  movel([-0.121105, -0.780827, -2.794142, -1.137419, 1.570796, 1.449692],accel_mss,speed_ms,0,blend_radius_m)
  movel([-0.120159, -0.781005, -2.794114, -1.137271, 1.570796, 1.450637],accel_mss,speed_ms,0,blend_radius_m)
  movel([-0.119008, -0.782524, -2.793869, -1.135997, 1.570796, 1.451789],accel_mss,speed_ms,0,blend_radius_m)
  movel([-0.118135, -0.785303, -2.793417, -1.133668, 1.570796, 1.452661],accel_mss,speed_ms,0,blend_radius_m)
  movel([-0.117601, -0.788380, -2.792913, -1.131096, 1.570796, 1.453195],accel_mss,speed_ms,0,blend_radius_m)
  movel([-0.115239, -0.783750, -2.793670, -1.134969, 1.570796, 1.455558],accel_mss,speed_ms,0,blend_radius_m)
  movel([-0.112520, -0.779061, -2.794425, -1.138903, 1.570796, 1.458276],accel_mss,speed_ms,0,blend_radius_m)
  movel([-0.109499, -0.774375, -2.795169, -1.142845, 1.570796, 1.461298],accel_mss,speed_ms,0,blend_radius_m)
  movel([-0.106241, -0.769762, -2.795890, -1.146737, 1.570796, 1.464556],accel_mss,speed_ms,0,blend_radius_m)
  movel([-0.099689, -0.760491, -2.797308, -1.154590, 1.570796, 1.471108],accel_mss,speed_ms,0,blend_radius_m)
  movel([-0.097728, -0.757937, -2.797692, -1.156760, 1.570796, 1.473068],accel_mss,speed_ms,0,blend_radius_m)
  movel([-0.095794, -0.755653, -2.798032, -1.158704, 1.570796, 1.475003],accel_mss,speed_ms,0,blend_radius_m)
  movel([-0.093954, -0.753818, -2.798303, -1.160268, 1.570796, 1.476842],accel_mss,speed_ms,0,blend_radius_m)
  movel([-0.092299, -0.752614, -2.798480, -1.161295, 1.570796, 1.478498],accel_mss,speed_ms,0,blend_radius_m)
  movel([-0.090884, -0.752253, -2.798533, -1.161603, 1.570796, 1.479912],accel_mss,speed_ms,0,blend_radius_m)
  movel([-0.089878, -0.752769, -2.798457, -1.161162, 1.570796, 1.480919],accel_mss,speed_ms,0,blend_radius_m)
  movel([-0.089251, -0.753972, -2.798280, -1.160137, 1.570796, 1.481545],accel_mss,speed_ms,0,blend_radius_m)
  movel([-0.088991, -0.755673, -2.798029, -1.158687, 1.570796, 1.481805],accel_mss,speed_ms,0,blend_radius_m)
  movel([-0.089073, -0.757680, -2.797730, -1.156979, 1.570796, 1.481724],accel_mss,speed_ms,0,blend_radius_m)
  movel([-0.089471, -0.759797, -2.797413, -1.155179, 1.570796, 1.481326],accel_mss,speed_ms,0,blend_radius_m)
  movel([-0.090165, -0.761839, -2.797105, -1.153445, 1.570796, 1.480631],accel_mss,speed_ms,0,blend_radius_m)
  movel([-0.091138, -0.763618, -2.796835, -1.151936, 1.570796, 1.479658],accel_mss,speed_ms,0,blend_radius_m)
  movel([-0.085055, -0.755408, -2.798068, -1.158913, 1.570796, 1.485742],accel_mss,speed_ms,0,blend_radius_m)
  movel([-0.081792, -0.751409, -2.798657, -1.162323, 1.570796, 1.489004],accel_mss,speed_ms,0,blend_radius_m)
  movel([-0.078396, -0.747530, -2.799220, -1.165639, 1.570796, 1.492400],accel_mss,speed_ms,0,blend_radius_m)
  movel([-0.074888, -0.743806, -2.799755, -1.168828, 1.570796, 1.495909],accel_mss,speed_ms,0,blend_radius_m)
  movel([-0.071275, -0.740275, -2.800255, -1.171859, 1.570796, 1.499521],accel_mss,speed_ms,0,blend_radius_m)
  movel([-0.067576, -0.736976, -2.800718, -1.174695, 1.570796, 1.503221],accel_mss,speed_ms,0,blend_radius_m)
  movel([-0.063806, -0.733944, -2.801138, -1.177307, 1.570796, 1.506991],accel_mss,speed_ms,0,blend_radius_m)
  movel([-0.061242, -0.732398, -2.801351, -1.178640, 1.570796, 1.509554],accel_mss,speed_ms,0,blend_radius_m)
  movel([-0.058496, -0.731434, -2.801483, -1.179472, 1.570796, 1.512301],accel_mss,speed_ms,0,blend_radius_m)
  movel([-0.057304, -0.731323, -2.801498, -1.179568, 1.570796, 1.513493],accel_mss,speed_ms,0,blend_radius_m)
  movel([-0.056360, -0.731534, -2.801469, -1.179386, 1.570796, 1.514437],accel_mss,speed_ms,0,blend_radius_m)
  movel([-0.055759, -0.732128, -2.801388, -1.178873, 1.570796, 1.515037],accel_mss,speed_ms,0,blend_radius_m)
  movel([-0.055607, -0.733168, -2.801245, -1.177976, 1.570796, 1.515190],accel_mss,speed_ms,0,blend_radius_m)
  movel([-0.055970, -0.734525, -2.801058, -1.176806, 1.570796, 1.514827],accel_mss,speed_ms,0,blend_radius_m)
  movel([-0.056714, -0.736045, -2.800847, -1.175497, 1.570796, 1.514083],accel_mss,speed_ms,0,blend_radius_m)
  movel([-0.058927, -0.739452, -2.800371, -1.172566, 1.570796, 1.511869],accel_mss,speed_ms,0,blend_radius_m)
  movel([-0.061573, -0.742637, -2.799921, -1.169831, 1.570796, 1.509223],accel_mss,speed_ms,0,blend_radius_m)
  movel([-0.064470, -0.745574, -2.799502, -1.167314, 1.570796, 1.506326],accel_mss,speed_ms,0,blend_radius_m)
  movel([-0.067437, -0.748234, -2.799119, -1.165036, 1.570796, 1.503359],accel_mss,speed_ms,0,blend_radius_m)
  movel([-0.063607, -0.746740, -2.799334, -1.166315, 1.570796, 1.507189],accel_mss,speed_ms,0,blend_radius_m)
  movel([-0.059620, -0.744795, -2.799614, -1.167981, 1.570796, 1.511176],accel_mss,speed_ms,0,blend_radius_m)
  movel([-0.055519, -0.742424, -2.799951, -1.170014, 1.570796, 1.515278],accel_mss,speed_ms,0,blend_radius_m)
  movel([-0.051338, -0.739647, -2.800344, -1.172398, 1.570796, 1.519459],accel_mss,speed_ms,0,blend_radius_m)
  movel([-0.048030, -0.737110, -2.800699, -1.174580, 1.570796, 1.522766],accel_mss,speed_ms,0,blend_radius_m)
  movel([-0.041537, -0.731618, -2.801458, -1.179314, 1.570796, 1.529259],accel_mss,speed_ms,0,blend_radius_m)
  movel([-0.038202, -0.729035, -2.801810, -1.181544, 1.570796, 1.532595],accel_mss,speed_ms,0,blend_radius_m)
  movel([-0.034400, -0.726366, -2.802170, -1.183853, 1.570796, 1.536396],accel_mss,speed_ms,0,blend_radius_m)
  movel([-0.027997, -0.722210, -2.802725, -1.187455, 1.570796, 1.542799],accel_mss,speed_ms,0,blend_radius_m)
  movel([-0.024935, -0.720489, -2.802952, -1.188948, 1.570796, 1.545861],accel_mss,speed_ms,0,blend_radius_m)
  movel([-0.022568, -0.719500, -2.803082, -1.189807, 1.570796, 1.548229],accel_mss,speed_ms,0,blend_radius_m)
  movel([-0.021784, -0.719391, -2.803096, -1.189901, 1.570796, 1.549013],accel_mss,speed_ms,0,blend_radius_m)
  movel([-0.021347, -0.719607, -2.803068, -1.189714, 1.570796, 1.549449],accel_mss,speed_ms,0,blend_radius_m)
  movel([-0.021306, -0.720180, -2.802993, -1.189216, 1.570796, 1.549490],accel_mss,speed_ms,0,blend_radius_m)
  movel([-0.021722, -0.721161, -2.802863, -1.188364, 1.570796, 1.549074],accel_mss,speed_ms,0,blend_radius_m)
  movel([-0.023301, -0.723619, -2.802538, -1.186232, 1.570796, 1.547495],accel_mss,speed_ms,0,blend_radius_m)
  movel([-0.025347, -0.726195, -2.802193, -1.184001, 1.570796, 1.545450],accel_mss,speed_ms,0,blend_radius_m)
  movel([-0.027725, -0.728828, -2.801838, -1.181723, 1.570796, 1.543072],accel_mss,speed_ms,0,blend_radius_m)
  movel([-0.030292, -0.731434, -2.801483, -1.179472, 1.570796, 1.540504],accel_mss,speed_ms,0,blend_radius_m)
  movel([-0.035478, -0.736292, -2.800813, -1.175284, 1.570796, 1.535318],accel_mss,speed_ms,0,blend_radius_m)
  movel([-0.039835, -0.740201, -2.800266, -1.171922, 1.570796, 1.530962],accel_mss,speed_ms,0,blend_radius_m)
  movel([-0.037640, -0.739808, -2.800321, -1.172260, 1.570796, 1.533156],accel_mss,speed_ms,0,blend_radius_m)
  movel([-0.035326, -0.739146, -2.800414, -1.172829, 1.570796, 1.535470],accel_mss,speed_ms,0,blend_radius_m)
  movel([-0.030418, -0.737158, -2.800692, -1.174539, 1.570796, 1.540378],accel_mss,speed_ms,0,blend_radius_m)
  movel([-0.025249, -0.734489, -2.801063, -1.176837, 1.570796, 1.545548],accel_mss,speed_ms,0,blend_radius_m)
  movel([-0.019955, -0.731399, -2.801488, -1.179502, 1.570796, 1.550841],accel_mss,speed_ms,0,blend_radius_m)
  movel([-0.015550, -0.728573, -2.801872, -1.181943, 1.570796, 1.555246],accel_mss,speed_ms,0,blend_radius_m)
  movel([-0.002182, -0.719511, -2.803081, -1.189798, 1.570796, 1.568614],accel_mss,speed_ms,0,blend_radius_m)
  movel([0.000291, -0.718246, -2.803246, -1.190897, 1.570796, 1.571087],accel_mss,speed_ms,0,blend_radius_m)
  movel([0.002219, -0.717829, -2.803301, -1.191260, 1.570796, 1.573015],accel_mss,speed_ms,0,blend_radius_m)
  movel([0.002614, -0.718141, -2.803260, -1.190988, 1.570796, 1.573410],accel_mss,speed_ms,0,blend_radius_m)
  movel([0.002432, -0.718911, -2.803159, -1.190319, 1.570796, 1.573228],accel_mss,speed_ms,0,blend_radius_m)
  movel([0.001528, -0.720216, -2.802988, -1.189185, 1.570796, 1.572325],accel_mss,speed_ms,0,blend_radius_m)
  movel([-0.000242, -0.722135, -2.802735, -1.187519, 1.570796, 1.570554],accel_mss,speed_ms,0,blend_radius_m)
  movel([-0.003204, -0.724919, -2.802364, -1.185106, 1.570796, 1.567592],accel_mss,speed_ms,0,blend_radius_m)
  movel([-0.006618, -0.727778, -2.801980, -1.182631, 1.570796, 1.564179],accel_mss,speed_ms,0,blend_radius_m)
  movel([-0.009977, -0.730186, -2.801653, -1.180550, 1.570796, 1.560819],accel_mss,speed_ms,0,blend_radius_m)
  movel([-0.011482, -0.731060, -2.801534, -1.179795, 1.570796, 1.559315],accel_mss,speed_ms,0,blend_radius_m)
  movel([-0.012779, -0.731617, -2.801458, -1.179315, 1.570796, 1.558017],accel_mss,speed_ms,0,blend_radius_m)
  movel([-0.007737, -0.731422, -2.801485, -1.179482, 1.570796, 1.563059],accel_mss,speed_ms,0,blend_radius_m)
  movel([-0.002332, -0.730537, -2.801605, -1.180246, 1.570796, 1.568464],accel_mss,speed_ms,0,blend_radius_m)
  movel([0.003362, -0.729092, -2.801802, -1.181495, 1.570796, 1.574158],accel_mss,speed_ms,0,blend_radius_m)
  movel([0.009278, -0.727224, -2.802055, -1.183111, 1.570796, 1.580074],accel_mss,speed_ms,0,blend_radius_m)
  movel([0.021466, -0.722735, -2.802655, -1.186999, 1.570796, 1.592262],accel_mss,speed_ms,0,blend_radius_m)
  movel([0.033600, -0.718155, -2.803258, -1.190976, 1.570796, 1.604396],accel_mss,speed_ms,0,blend_radius_m)
  movel([0.035605, -0.717735, -2.803313, -1.191341, 1.570796, 1.606402],accel_mss,speed_ms,0,blend_radius_m)
  movel([0.036255, -0.718010, -2.803277, -1.191101, 1.570796, 1.607051],accel_mss,speed_ms,0,blend_radius_m)
  movel([0.036422, -0.718815, -2.803172, -1.190402, 1.570796, 1.607218],accel_mss,speed_ms,0,blend_radius_m)
  movel([0.036036, -0.720000, -2.803016, -1.189373, 1.570796, 1.606833],accel_mss,speed_ms,0,blend_radius_m)
  movel([0.034004, -0.723279, -2.802583, -1.186527, 1.570796, 1.604800],accel_mss,speed_ms,0,blend_radius_m)
  movel([0.032557, -0.725161, -2.802332, -1.184896, 1.570796, 1.603354],accel_mss,speed_ms,0,blend_radius_m)
  movel([0.029315, -0.728658, -2.801861, -1.181870, 1.570796, 1.600111],accel_mss,speed_ms,0,blend_radius_m)
  movel([0.025758, -0.731771, -2.801437, -1.179181, 1.570796, 1.596555],accel_mss,speed_ms,0,blend_radius_m)
  movel([0.022037, -0.734500, -2.801061, -1.176828, 1.570796, 1.592834],accel_mss,speed_ms,0,blend_radius_m)
  movel([0.018315, -0.736820, -2.800739, -1.174829, 1.570796, 1.589112],accel_mss,speed_ms,0,blend_radius_m)
  movel([0.014745, -0.738726, -2.800473, -1.173190, 1.570796, 1.585541],accel_mss,speed_ms,0,blend_radius_m)
  movel([0.011481, -0.740197, -2.800266, -1.171925, 1.570796, 1.582277],accel_mss,speed_ms,0,blend_radius_m)
  movel([0.008687, -0.741208, -2.800124, -1.171057, 1.570796, 1.579483],accel_mss,speed_ms,0,blend_radius_m)
  movel([0.008653, -0.742047, -2.800005, -1.170337, 1.570796, 1.579449],accel_mss,speed_ms,0,blend_radius_m)
  movel([0.009139, -0.742448, -2.799948, -1.169993, 1.570796, 1.579935],accel_mss,speed_ms,0,blend_radius_m)
  movel([0.010647, -0.742839, -2.799892, -1.169658, 1.570796, 1.581444],accel_mss,speed_ms,0,blend_radius_m)
  movel([0.012360, -0.742904, -2.799883, -1.169602, 1.570796, 1.583157],accel_mss,speed_ms,0,blend_radius_m)
  movel([0.016128, -0.742457, -2.799947, -1.169986, 1.570796, 1.586925],accel_mss,speed_ms,0,blend_radius_m)
  movel([0.022850, -0.741236, -2.800120, -1.171033, 1.570796, 1.593647],accel_mss,speed_ms,0,blend_radius_m)
  movel([0.029687, -0.739729, -2.800332, -1.172328, 1.570796, 1.600483],accel_mss,speed_ms,0,blend_radius_m)
  movel([0.043712, -0.735971, -2.800858, -1.175560, 1.570796, 1.614508],accel_mss,speed_ms,0,blend_radius_m)
  movel([0.047601, -0.735012, -2.800990, -1.176386, 1.570796, 1.618397],accel_mss,speed_ms,0,blend_radius_m)
  movel([0.050057, -0.734636, -2.801043, -1.176710, 1.570796, 1.620854],accel_mss,speed_ms,0,blend_radius_m)
  movel([0.052405, -0.734564, -2.801053, -1.176772, 1.570796, 1.623201],accel_mss,speed_ms,0,blend_radius_m)
  movel([0.054288, -0.734979, -2.800995, -1.176415, 1.570796, 1.625084],accel_mss,speed_ms,0,blend_radius_m)
  movel([0.055366, -0.736045, -2.800847, -1.175497, 1.570796, 1.626162],accel_mss,speed_ms,0,blend_radius_m)
  movel([0.055503, -0.736869, -2.800733, -1.174788, 1.570796, 1.626300],accel_mss,speed_ms,0,blend_radius_m)
  movel([0.055317, -0.737917, -2.800586, -1.173885, 1.570796, 1.626113],accel_mss,speed_ms,0,blend_radius_m)
  movel([0.054755, -0.739218, -2.800404, -1.172767, 1.570796, 1.625552],accel_mss,speed_ms,0,blend_radius_m)
  movel([0.053791, -0.740777, -2.800184, -1.171427, 1.570796, 1.624588],accel_mss,speed_ms,0,blend_radius_m)
  movel([0.052380, -0.742206, -2.799982, -1.170200, 1.570796, 1.623176],accel_mss,speed_ms,0,blend_radius_m)
  movel([0.050460, -0.743557, -2.799790, -1.169042, 1.570796, 1.621256],accel_mss,speed_ms,0,blend_radius_m)
  movel([0.040183, -0.749654, -2.798913, -1.163823, 1.570796, 1.610979],accel_mss,speed_ms,0,blend_radius_m)
  movel([0.036738, -0.751253, -2.798679, -1.162457, 1.570796, 1.607535],accel_mss,speed_ms,0,blend_radius_m)
  movel([0.035260, -0.751698, -2.798614, -1.162077, 1.570796, 1.606056],accel_mss,speed_ms,0,blend_radius_m)
  movel([0.034042, -0.751799, -2.798600, -1.161990, 1.570796, 1.604838],accel_mss,speed_ms,0,blend_radius_m)
  movel([0.039097, -0.753329, -2.798375, -1.160685, 1.570796, 1.609893],accel_mss,speed_ms,0,blend_radius_m)
  movel([0.044720, -0.753966, -2.798281, -1.160142, 1.570796, 1.615516],accel_mss,speed_ms,0,blend_radius_m)
  movel([0.050778, -0.753874, -2.798295, -1.160221, 1.570796, 1.621574],accel_mss,speed_ms,0,blend_radius_m)
  movel([0.057144, -0.753204, -2.798393, -1.160792, 1.570796, 1.627940],accel_mss,speed_ms,0,blend_radius_m)
  movel([0.062648, -0.751826, -2.798596, -1.161967, 1.570796, 1.633444],accel_mss,speed_ms,0,blend_radius_m)
  movel([0.070534, -0.750016, -2.798860, -1.163513, 1.570796, 1.641330],accel_mss,speed_ms,0,blend_radius_m)
  movel([0.074102, -0.749639, -2.798915, -1.163835, 1.570796, 1.644899],accel_mss,speed_ms,0,blend_radius_m)
  movel([0.076754, -0.749965, -2.798867, -1.163557, 1.570796, 1.647550],accel_mss,speed_ms,0,blend_radius_m)
  movel([0.077577, -0.750472, -2.798793, -1.163123, 1.570796, 1.648374],accel_mss,speed_ms,0,blend_radius_m)
  movel([0.077981, -0.751251, -2.798680, -1.162459, 1.570796, 1.648777],accel_mss,speed_ms,0,blend_radius_m)
  movel([0.077904, -0.752336, -2.798521, -1.161532, 1.570796, 1.648701],accel_mss,speed_ms,0,blend_radius_m)
  movel([0.077296, -0.753748, -2.798313, -1.160328, 1.570796, 1.648093],accel_mss,speed_ms,0,blend_radius_m)
  movel([0.076368, -0.755193, -2.798100, -1.159096, 1.570796, 1.647164],accel_mss,speed_ms,0,blend_radius_m)
  movel([0.075295, -0.756570, -2.797895, -1.157924, 1.570796, 1.646091],accel_mss,speed_ms,0,blend_radius_m)
  movel([0.072924, -0.759131, -2.797513, -1.155746, 1.570796, 1.643720],accel_mss,speed_ms,0,blend_radius_m)
  movel([0.070302, -0.761655, -2.797133, -1.153602, 1.570796, 1.641099],accel_mss,speed_ms,0,blend_radius_m)
  movel([0.064988, -0.766133, -2.796451, -1.149806, 1.570796, 1.635784],accel_mss,speed_ms,0,blend_radius_m)
  movel([0.062326, -0.768067, -2.796153, -1.148169, 1.570796, 1.633122],accel_mss,speed_ms,0,blend_radius_m)
  movel([0.067181, -0.767478, -2.796244, -1.148667, 1.570796, 1.637977],accel_mss,speed_ms,0,blend_radius_m)
  movel([0.072189, -0.766515, -2.796392, -1.149482, 1.570796, 1.642985],accel_mss,speed_ms,0,blend_radius_m)
  movel([0.077338, -0.765224, -2.796590, -1.150576, 1.570796, 1.648134],accel_mss,speed_ms,0,blend_radius_m)
  movel([0.082615, -0.763635, -2.796832, -1.151922, 1.570796, 1.653412],accel_mss,speed_ms,0,blend_radius_m)
  movel([0.093490, -0.759739, -2.797422, -1.155229, 1.570796, 1.664286],accel_mss,speed_ms,0,blend_radius_m)
  movel([0.104701, -0.755125, -2.798110, -1.159154, 1.570796, 1.675497],accel_mss,speed_ms,0,blend_radius_m)
  movel([0.107639, -0.754225, -2.798243, -1.159921, 1.570796, 1.678435],accel_mss,speed_ms,0,blend_radius_m)
  movel([0.108683, -0.754415, -2.798215, -1.159759, 1.570796, 1.679480],accel_mss,speed_ms,0,blend_radius_m)
  movel([0.109107, -0.755353, -2.798076, -1.158960, 1.570796, 1.679903],accel_mss,speed_ms,0,blend_radius_m)
  movel([0.108974, -0.756313, -2.797934, -1.158142, 1.570796, 1.679770],accel_mss,speed_ms,0,blend_radius_m)
  movel([0.108569, -0.757391, -2.797773, -1.157225, 1.570796, 1.679365],accel_mss,speed_ms,0,blend_radius_m)
  movel([0.107060, -0.759842, -2.797406, -1.155141, 1.570796, 1.677856],accel_mss,speed_ms,0,blend_radius_m)
  movel([0.104857, -0.762515, -2.797002, -1.152872, 1.570796, 1.675653],accel_mss,speed_ms,0,blend_radius_m)
  movel([0.102226, -0.765245, -2.796587, -1.150558, 1.570796, 1.673022],accel_mss,speed_ms,0,blend_radius_m)
  movel([0.096762, -0.770165, -2.795828, -1.146396, 1.570796, 1.667558],accel_mss,speed_ms,0,blend_radius_m)
  movel([0.092780, -0.773214, -2.795351, -1.143823, 1.570796, 1.663577],accel_mss,speed_ms,0,blend_radius_m)
  movel([0.095018, -0.772547, -2.795456, -1.144386, 1.570796, 1.665815],accel_mss,speed_ms,0,blend_radius_m)
  movel([0.097342, -0.771623, -2.795601, -1.145166, 1.570796, 1.668138],accel_mss,speed_ms,0,blend_radius_m)
  movel([0.102193, -0.769088, -2.795995, -1.147306, 1.570796, 1.672990],accel_mss,speed_ms,0,blend_radius_m)
  movel([0.107238, -0.765717, -2.796514, -1.150158, 1.570796, 1.678035],accel_mss,speed_ms,0,blend_radius_m)
  movel([0.112383, -0.761637, -2.797135, -1.153617, 1.570796, 1.683179],accel_mss,speed_ms,0,blend_radius_m)
  movel([0.117534, -0.756944, -2.797840, -1.157606, 1.570796, 1.688330],accel_mss,speed_ms,0,blend_radius_m)
  movel([0.122590, -0.751769, -2.798604, -1.162016, 1.570796, 1.693387],accel_mss,speed_ms,0,blend_radius_m)
  movel([0.127452, -0.746216, -2.799410, -1.166763, 1.570796, 1.698249],accel_mss,speed_ms,0,blend_radius_m)
  movel([0.132018, -0.740413, -2.800236, -1.171740, 1.570796, 1.702814],accel_mss,speed_ms,0,blend_radius_m)
  movel([0.134037, -0.737820, -2.800600, -1.173969, 1.570796, 1.704834],accel_mss,speed_ms,0,blend_radius_m)
  movel([0.135120, -0.736689, -2.800758, -1.174942, 1.570796, 1.705916],accel_mss,speed_ms,0,blend_radius_m)
  movel([0.136237, -0.735818, -2.800879, -1.175692, 1.570796, 1.707033],accel_mss,speed_ms,0,blend_radius_m)
  movel([0.137379, -0.735340, -2.800945, -1.176104, 1.570796, 1.708175],accel_mss,speed_ms,0,blend_radius_m)
  movel([0.138333, -0.735302, -2.800950, -1.176136, 1.570796, 1.709129],accel_mss,speed_ms,0,blend_radius_m)
  movel([0.139345, -0.735960, -2.800859, -1.175570, 1.570796, 1.710141],accel_mss,speed_ms,0,blend_radius_m)
  movel([0.139829, -0.737373, -2.800662, -1.174353, 1.570796, 1.710625],accel_mss,speed_ms,0,blend_radius_m)
  movel([0.139879, -0.739349, -2.800386, -1.172654, 1.570796, 1.710675],accel_mss,speed_ms,0,blend_radius_m)
  movel([0.139591, -0.741712, -2.800052, -1.170625, 1.570796, 1.710387],accel_mss,speed_ms,0,blend_radius_m)
  movel([0.138373, -0.746843, -2.799319, -1.166227, 1.570796, 1.709169],accel_mss,speed_ms,0,blend_radius_m)
  movel([0.136926, -0.751311, -2.798671, -1.162407, 1.570796, 1.707723],accel_mss,speed_ms,0,blend_radius_m)
  movel([0.140852, -0.745658, -2.799490, -1.167241, 1.570796, 1.711648],accel_mss,speed_ms,0,blend_radius_m)
  movel([0.144402, -0.739896, -2.800309, -1.172184, 1.570796, 1.715198],accel_mss,speed_ms,0,blend_radius_m)
  movel([0.147549, -0.734083, -2.801119, -1.177187, 1.570796, 1.718345],accel_mss,speed_ms,0,blend_radius_m)
  movel([0.150273, -0.728298, -2.801910, -1.182182, 1.570796, 1.721070],accel_mss,speed_ms,0,blend_radius_m)
  movel([0.152533, -0.722617, -2.802671, -1.187101, 1.570796, 1.723330],accel_mss,speed_ms,0,blend_radius_m)
  movel([0.154318, -0.717103, -2.803395, -1.191890, 1.570796, 1.725114],accel_mss,speed_ms,0,blend_radius_m)
  movel([0.155580, -0.711854, -2.804072, -1.196463, 1.570796, 1.726376],accel_mss,speed_ms,0,blend_radius_m)
  movel([0.156297, -0.706938, -2.804695, -1.200756, 1.570796, 1.727094],accel_mss,speed_ms,0,blend_radius_m)
  movel([0.156402, -0.700717, -2.805467, -1.206205, 1.570796, 1.727198],accel_mss,speed_ms,0,blend_radius_m)
  movel([0.156716, -0.697272, -2.805887, -1.209229, 1.570796, 1.727512],accel_mss,speed_ms,0,blend_radius_m)
  movel([0.157110, -0.695510, -2.806100, -1.210779, 1.570796, 1.727906],accel_mss,speed_ms,0,blend_radius_m)
  movel([0.157721, -0.693740, -2.806313, -1.212336, 1.570796, 1.728517],accel_mss,speed_ms,0,blend_radius_m)
  movel([0.159157, -0.690828, -2.806659, -1.214902, 1.570796, 1.729953],accel_mss,speed_ms,0,blend_radius_m)
  movel([0.160486, -0.689041, -2.806870, -1.216478, 1.570796, 1.731283],accel_mss,speed_ms,0,blend_radius_m)
  movel([0.161725, -0.688141, -2.806976, -1.217273, 1.570796, 1.732521],accel_mss,speed_ms,0,blend_radius_m)
  movel([0.162880, -0.687888, -2.807005, -1.217496, 1.570796, 1.733676],accel_mss,speed_ms,0,blend_radius_m)
  movel([0.165920, -0.688642, -2.806917, -1.216830, 1.570796, 1.736716],accel_mss,speed_ms,0,blend_radius_m)
  movel([0.166833, -0.688590, -2.806923, -1.216876, 1.570796, 1.737629],accel_mss,speed_ms,0,blend_radius_m)
  movel([0.168876, -0.684269, -2.807426, -1.220694, 1.570796, 1.739672],accel_mss,speed_ms,0,blend_radius_m)
  movel([0.170617, -0.679986, -2.807917, -1.224486, 1.570796, 1.741413],accel_mss,speed_ms,0,blend_radius_m)
  movel([0.172069, -0.675763, -2.808393, -1.228233, 1.570796, 1.742866],accel_mss,speed_ms,0,blend_radius_m)
  movel([0.173248, -0.671607, -2.808854, -1.231928, 1.570796, 1.744044],accel_mss,speed_ms,0,blend_radius_m)
  movel([0.174153, -0.667546, -2.809297, -1.235545, 1.570796, 1.744950],accel_mss,speed_ms,0,blend_radius_m)
  movel([0.174801, -0.663592, -2.809722, -1.239075, 1.570796, 1.745598],accel_mss,speed_ms,0,blend_radius_m)
  movel([0.175391, -0.656055, -2.810514, -1.245820, 1.570796, 1.746188],accel_mss,speed_ms,0,blend_radius_m)
  movel([0.175103, -0.649147, -2.811218, -1.252023, 1.570796, 1.745899],accel_mss,speed_ms,0,blend_radius_m)
  movel([0.174059, -0.642982, -2.811830, -1.257577, 1.570796, 1.744855],accel_mss,speed_ms,0,blend_radius_m)
  movel([0.172351, -0.637702, -2.812342, -1.262345, 1.570796, 1.743147],accel_mss,speed_ms,0,blend_radius_m)
  movel([0.170116, -0.633411, -2.812749, -1.266228, 1.570796, 1.740912],accel_mss,speed_ms,0,blend_radius_m)
  speed_ms = 0.005
  movel([0.170116, -0.627529, -2.805977, -1.278883, 1.570796, 1.740912],accel_mss,speed_ms,0,blend_radius_m)
  speed_ms = 0.040
  movel([0.138700, -0.651920, -2.803568, -1.256901, 1.570796, 1.709497],accel_mss,speed_ms,0,blend_radius_m)
  speed_ms = 0.005
  movel([0.138700, -0.658181, -2.810293, -1.243915, 1.570796, 1.709497],accel_mss,speed_ms,0,blend_radius_m)
  speed_ms = 0.025
  movel([0.136102, -0.657818, -2.810331, -1.244240, 1.570796, 1.706899],accel_mss,speed_ms,0,blend_radius_m)
  movel([0.133054, -0.658341, -2.810276, -1.243772, 1.570796, 1.703850],accel_mss,speed_ms,0,blend_radius_m)
  movel([0.129644, -0.659620, -2.810142, -1.242627, 1.570796, 1.700441],accel_mss,speed_ms,0,blend_radius_m)
  movel([0.125976, -0.661510, -2.809943, -1.240936, 1.570796, 1.696772],accel_mss,speed_ms,0,blend_radius_m)
  movel([0.122143, -0.663876, -2.809692, -1.238821, 1.570796, 1.692939],accel_mss,speed_ms,0,blend_radius_m)
  movel([0.118234, -0.666581, -2.809402, -1.236407, 1.570796, 1.689030],accel_mss,speed_ms,0,blend_radius_m)
  movel([0.110564, -0.672460, -2.808760, -1.231169, 1.570796, 1.681360],accel_mss,speed_ms,0,blend_radius_m)
  speed_ms = 0.005
  movel([0.110564, -0.665989, -2.802064, -1.244335, 1.570796, 1.681360],accel_mss,speed_ms,0,blend_radius_m)
  speed_ms = 0.040
  movel([0.120496, -0.657640, -2.802967, -1.251782, 1.570796, 1.691293],accel_mss,speed_ms,0,blend_radius_m)
  speed_ms = 0.005
  movel([0.120496, -0.663987, -2.809680, -1.238722, 1.570796, 1.691293],accel_mss,speed_ms,0,blend_radius_m)
  speed_ms = 0.025
  movel([0.122110, -0.659259, -2.810180, -1.242950, 1.570796, 1.692907],accel_mss,speed_ms,0,blend_radius_m)
  movel([0.123299, -0.654866, -2.810636, -1.246887, 1.570796, 1.694095],accel_mss,speed_ms,0,blend_radius_m)
  movel([0.124068, -0.650800, -2.811051, -1.250538, 1.570796, 1.694864],accel_mss,speed_ms,0,blend_radius_m)
  movel([0.124435, -0.647046, -2.811429, -1.253915, 1.570796, 1.695231],accel_mss,speed_ms,0,blend_radius_m)
  movel([0.124423, -0.643584, -2.811771, -1.257034, 1.570796, 1.695219],accel_mss,speed_ms,0,blend_radius_m)
  movel([0.124046, -0.640402, -2.812082, -1.259905, 1.570796, 1.694842],accel_mss,speed_ms,0,blend_radius_m)
  movel([0.123323, -0.637484, -2.812363, -1.262542, 1.570796, 1.694119],accel_mss,speed_ms,0,blend_radius_m)
  movel([0.122274, -0.634812, -2.812617, -1.264960, 1.570796, 1.693071],accel_mss,speed_ms,0,blend_radius_m)
  movel([0.118229, -0.627978, -2.813255, -1.271156, 1.570796, 1.689025],accel_mss,speed_ms,0,blend_radius_m)
  movel([0.116481, -0.624510, -2.813571, -1.274308, 1.570796, 1.687277],accel_mss,speed_ms,0,blend_radius_m)
  movel([0.115290, -0.620006, -2.813974, -1.278409, 1.570796, 1.686086],accel_mss,speed_ms,0,blend_radius_m)
  movel([0.114590, -0.613627, -2.814532, -1.284231, 1.570796, 1.685386],accel_mss,speed_ms,0,blend_radius_m)
  movel([0.114549, -0.606649, -2.815123, -1.290617, 1.570796, 1.685345],accel_mss,speed_ms,0,blend_radius_m)
  movel([0.115398, -0.598953, -2.815753, -1.297683, 1.570796, 1.686195],accel_mss,speed_ms,0,blend_radius_m)
  movel([0.116229, -0.594796, -2.816083, -1.301510, 1.570796, 1.687025],accel_mss,speed_ms,0,blend_radius_m)
  movel([0.117376, -0.590413, -2.816425, -1.305551, 1.570796, 1.688172],accel_mss,speed_ms,0,blend_radius_m)
  movel([0.119840, -0.583271, -2.816965, -1.312154, 1.570796, 1.690636],accel_mss,speed_ms,0,blend_radius_m)
  movel([0.123098, -0.575926, -2.817500, -1.318963, 1.570796, 1.693894],accel_mss,speed_ms,0,blend_radius_m)
  movel([0.127112, -0.568433, -2.818025, -1.325932, 1.570796, 1.697908],accel_mss,speed_ms,0,blend_radius_m)
  movel([0.131842, -0.560852, -2.818534, -1.333004, 1.570796, 1.702638],accel_mss,speed_ms,0,blend_radius_m)
  movel([0.137234, -0.553260, -2.819022, -1.340107, 1.570796, 1.708030],accel_mss,speed_ms,0,blend_radius_m)
  movel([0.143247, -0.545723, -2.819486, -1.347180, 1.570796, 1.714044],accel_mss,speed_ms,0,blend_radius_m)
  movel([0.149829, -0.538311, -2.819921, -1.354157, 1.570796, 1.720625],accel_mss,speed_ms,0,blend_radius_m)
  movel([0.156913, -0.531114, -2.820325, -1.360951, 1.570796, 1.727709],accel_mss,speed_ms,0,blend_radius_m)
  movel([0.162439, -0.525991, -2.820600, -1.365798, 1.570796, 1.733235],accel_mss,speed_ms,0,blend_radius_m)
  movel([0.168059, -0.521192, -2.820850, -1.370347, 1.570796, 1.738855],accel_mss,speed_ms,0,blend_radius_m)
  movel([0.173713, -0.516760, -2.821073, -1.374556, 1.570796, 1.744510],accel_mss,speed_ms,0,blend_radius_m)
  movel([0.179359, -0.512711, -2.821271, -1.378407, 1.570796, 1.750155],accel_mss,speed_ms,0,blend_radius_m)
  movel([0.184932, -0.509099, -2.821442, -1.381848, 1.570796, 1.755728],accel_mss,speed_ms,0,blend_radius_m)
  movel([0.190379, -0.505951, -2.821587, -1.384851, 1.570796, 1.761175],accel_mss,speed_ms,0,blend_radius_m)
  movel([0.195640, -0.503301, -2.821707, -1.387381, 1.570796, 1.766437],accel_mss,speed_ms,0,blend_radius_m)
  movel([0.200660, -0.501187, -2.821801, -1.389401, 1.570796, 1.771456],accel_mss,speed_ms,0,blend_radius_m)
  movel([0.205378, -0.499641, -2.821868, -1.390880, 1.570796, 1.776175],accel_mss,speed_ms,0,blend_radius_m)
  movel([0.209750, -0.498684, -2.821910, -1.391795, 1.570796, 1.780546],accel_mss,speed_ms,0,blend_radius_m)
  movel([0.213716, -0.498354, -2.821924, -1.392111, 1.570796, 1.784512],accel_mss,speed_ms,0,blend_radius_m)
  movel([0.217226, -0.498672, -2.821910, -1.391806, 1.570796, 1.788023],accel_mss,speed_ms,0,blend_radius_m)
  movel([0.220235, -0.499660, -2.821868, -1.390861, 1.570796, 1.791031],accel_mss,speed_ms,0,blend_radius_m)
  movel([0.222682, -0.501351, -2.821794, -1.389244, 1.570796, 1.793478],accel_mss,speed_ms,0,blend_radius_m)
  movel([0.224532, -0.503750, -2.821687, -1.386952, 1.570796, 1.795329],accel_mss,speed_ms,0,blend_radius_m)
  movel([0.225745, -0.506882, -2.821545, -1.383962, 1.570796, 1.796541],accel_mss,speed_ms,0,blend_radius_m)
  movel([0.226531, -0.511750, -2.821317, -1.379322, 1.570796, 1.797328],accel_mss,speed_ms,0,blend_radius_m)
  movel([0.226728, -0.517163, -2.821053, -1.374173, 1.570796, 1.797524],accel_mss,speed_ms,0,blend_radius_m)
  movel([0.226455, -0.522993, -2.820757, -1.368639, 1.570796, 1.797251],accel_mss,speed_ms,0,blend_radius_m)
  movel([0.225856, -0.529082, -2.820435, -1.362871, 1.570796, 1.796653],accel_mss,speed_ms,0,blend_radius_m)
  movel([0.223911, -0.542770, -2.819662, -1.349958, 1.570796, 1.794707],accel_mss,speed_ms,0,blend_radius_m)
  movel([0.221348, -0.556882, -2.818792, -1.336715, 1.570796, 1.792145],accel_mss,speed_ms,0,blend_radius_m)
  movel([0.218336, -0.571276, -2.817828, -1.323285, 1.570796, 1.789132],accel_mss,speed_ms,0,blend_radius_m)
  movel([0.215033, -0.585792, -2.816776, -1.309821, 1.570796, 1.785830],accel_mss,speed_ms,0,blend_radius_m)
  movel([0.201838, -0.642595, -2.811868, -1.257926, 1.570796, 1.772635],accel_mss,speed_ms,0,blend_radius_m)
  movel([0.196552, -0.669300, -2.809107, -1.233983, 1.570796, 1.767348],accel_mss,speed_ms,0,blend_radius_m)
  movel([0.194383, -0.682184, -2.807666, -1.222539, 1.570796, 1.765179],accel_mss,speed_ms,0,blend_radius_m)
  movel([0.192649, -0.694648, -2.806204, -1.211537, 1.570796, 1.763445],accel_mss,speed_ms,0,blend_radius_m)
  movel([0.191422, -0.706638, -2.804733, -1.201018, 1.570796, 1.762219],accel_mss,speed_ms,0,blend_radius_m)
  movel([0.190783, -0.718085, -2.803267, -1.191036, 1.570796, 1.761579],accel_mss,speed_ms,0,blend_radius_m)
  movel([0.190794, -0.728945, -2.801822, -1.181622, 1.570796, 1.761590],accel_mss,speed_ms,0,blend_radius_m)
  movel([0.191537, -0.739159, -2.800412, -1.172818, 1.570796, 1.762333],accel_mss,speed_ms,0,blend_radius_m)
  movel([0.192118, -0.742879, -2.799887, -1.169623, 1.570796, 1.762914],accel_mss,speed_ms,0,blend_radius_m)
  movel([0.193186, -0.746130, -2.799422, -1.166837, 1.570796, 1.763982],accel_mss,speed_ms,0,blend_radius_m)
  movel([0.194999, -0.748474, -2.799084, -1.164831, 1.570796, 1.765795],accel_mss,speed_ms,0,blend_radius_m)
  movel([0.196267, -0.749168, -2.798983, -1.164237, 1.570796, 1.767064],accel_mss,speed_ms,0,blend_radius_m)
  movel([0.197826, -0.749467, -2.798940, -1.163982, 1.570796, 1.768623],accel_mss,speed_ms,0,blend_radius_m)
  speed_ms = 0.005
  movel([0.197826, -0.741971, -2.792425, -1.177993, 1.570796, 1.768623],accel_mss,speed_ms,0,blend_radius_m)
  speed_ms = 0.040
  movel([0.166317, -0.704429, -2.797516, -1.210444, 1.570796, 1.737113],accel_mss,speed_ms,0,blend_radius_m)
  speed_ms = 0.005
  movel([0.166317, -0.711442, -2.804125, -1.196822, 1.570796, 1.737113],accel_mss,speed_ms,0,blend_radius_m)
  speed_ms = 0.025
  movel([0.165098, -0.713361, -2.803879, -1.195149, 1.570796, 1.735894],accel_mss,speed_ms,0,blend_radius_m)
  movel([0.164169, -0.715319, -2.803627, -1.193443, 1.570796, 1.734965],accel_mss,speed_ms,0,blend_radius_m)
  movel([0.163511, -0.717289, -2.803371, -1.191729, 1.570796, 1.734307],accel_mss,speed_ms,0,blend_radius_m)
  movel([0.163074, -0.719282, -2.803111, -1.189996, 1.570796, 1.733870],accel_mss,speed_ms,0,blend_radius_m)
  movel([0.162764, -0.723266, -2.802585, -1.186538, 1.570796, 1.733560],accel_mss,speed_ms,0,blend_radius_m)
  movel([0.162975, -0.727201, -2.802058, -1.183131, 1.570796, 1.733771],accel_mss,speed_ms,0,blend_radius_m)
  movel([0.164204, -0.737962, -2.800580, -1.173847, 1.570796, 1.735001],accel_mss,speed_ms,0,blend_radius_m)
  movel([0.163980, -0.740945, -2.800161, -1.171283, 1.570796, 1.734776],accel_mss,speed_ms,0,blend_radius_m)
  movel([0.163462, -0.742430, -2.799950, -1.170008, 1.570796, 1.734258],accel_mss,speed_ms,0,blend_radius_m)
  movel([0.162572, -0.743702, -2.799770, -1.168918, 1.570796, 1.733369],accel_mss,speed_ms,0,blend_radius_m)
  movel([0.161731, -0.744465, -2.799661, -1.168263, 1.570796, 1.732527],accel_mss,speed_ms,0,blend_radius_m)
  movel([0.160936, -0.744777, -2.799616, -1.167996, 1.570796, 1.731733],accel_mss,speed_ms,0,blend_radius_m)
  movel([0.160186, -0.744702, -2.799627, -1.168060, 1.570796, 1.730982],accel_mss,speed_ms,0,blend_radius_m)
  movel([0.158834, -0.743593, -2.799785, -1.169010, 1.570796, 1.729630],accel_mss,speed_ms,0,blend_radius_m)
  movel([0.157687, -0.741595, -2.800069, -1.170725, 1.570796, 1.728483],accel_mss,speed_ms,0,blend_radius_m)
  movel([0.156071, -0.736709, -2.800755, -1.174925, 1.570796, 1.726867],accel_mss,speed_ms,0,blend_radius_m)
  movel([0.155517, -0.733612, -2.801184, -1.177593, 1.570796, 1.726314],accel_mss,speed_ms,0,blend_radius_m)
  movel([0.153840, -0.739175, -2.800410, -1.172804, 1.570796, 1.724636],accel_mss,speed_ms,0,blend_radius_m)
  movel([0.152864, -0.744357, -2.799676, -1.168356, 1.570796, 1.723661],accel_mss,speed_ms,0,blend_radius_m)
  movel([0.152485, -0.749189, -2.798980, -1.164220, 1.570796, 1.723281],accel_mss,speed_ms,0,blend_radius_m)
  movel([0.152612, -0.753673, -2.798324, -1.160391, 1.570796, 1.723409],accel_mss,speed_ms,0,blend_radius_m)
  movel([0.153139, -0.757847, -2.797705, -1.156837, 1.570796, 1.723935],accel_mss,speed_ms,0,blend_radius_m)
  movel([0.153986, -0.761708, -2.797125, -1.153556, 1.570796, 1.724782],accel_mss,speed_ms,0,blend_radius_m)
  movel([0.156246, -0.768568, -2.796075, -1.147746, 1.570796, 1.727042],accel_mss,speed_ms,0,blend_radius_m)
  movel([0.156304, -0.770203, -2.795822, -1.146364, 1.570796, 1.727100],accel_mss,speed_ms,0,blend_radius_m)
  movel([0.155931, -0.771134, -2.795677, -1.145578, 1.570796, 1.726728],accel_mss,speed_ms,0,blend_radius_m)
  movel([0.155223, -0.771923, -2.795554, -1.144912, 1.570796, 1.726019],accel_mss,speed_ms,0,blend_radius_m)
  movel([0.154317, -0.772303, -2.795494, -1.144592, 1.570796, 1.725113],accel_mss,speed_ms,0,blend_radius_m)
  movel([0.152367, -0.772470, -2.795468, -1.144451, 1.570796, 1.723163],accel_mss,speed_ms,0,blend_radius_m)
  movel([0.150735, -0.772134, -2.795521, -1.144734, 1.570796, 1.721532],accel_mss,speed_ms,0,blend_radius_m)
  movel([0.149384, -0.771372, -2.795640, -1.145377, 1.570796, 1.720180],accel_mss,speed_ms,0,blend_radius_m)
  movel([0.148290, -0.770236, -2.795817, -1.146336, 1.570796, 1.719086],accel_mss,speed_ms,0,blend_radius_m)
  movel([0.146758, -0.767125, -2.796298, -1.148966, 1.570796, 1.717554],accel_mss,speed_ms,0,blend_radius_m)
  movel([0.145914, -0.763325, -2.796879, -1.152185, 1.570796, 1.716710],accel_mss,speed_ms,0,blend_radius_m)
  movel([0.145148, -0.772058, -2.795533, -1.144799, 1.570796, 1.715944],accel_mss,speed_ms,0,blend_radius_m)
  movel([0.145196, -0.776055, -2.794904, -1.141430, 1.570796, 1.715993],accel_mss,speed_ms,0,blend_radius_m)
  movel([0.145776, -0.779640, -2.794333, -1.138417, 1.570796, 1.716573],accel_mss,speed_ms,0,blend_radius_m)
  movel([0.146955, -0.782146, -2.793930, -1.136314, 1.570796, 1.717752],accel_mss,speed_ms,0,blend_radius_m)
  movel([0.150125, -0.785983, -2.793306, -1.133099, 1.570796, 1.720921],accel_mss,speed_ms,0,blend_radius_m)
  movel([0.151210, -0.788468, -2.792899, -1.131022, 1.570796, 1.722006],accel_mss,speed_ms,0,blend_radius_m)
  movel([0.151294, -0.789089, -2.792796, -1.130504, 1.570796, 1.722090],accel_mss,speed_ms,0,blend_radius_m)
  movel([0.151105, -0.789869, -2.792667, -1.129852, 1.570796, 1.721902],accel_mss,speed_ms,0,blend_radius_m)
  movel([0.150490, -0.790703, -2.792529, -1.129156, 1.570796, 1.721287],accel_mss,speed_ms,0,blend_radius_m)
  movel([0.149467, -0.791500, -2.792397, -1.128492, 1.570796, 1.720263],accel_mss,speed_ms,0,blend_radius_m)
  movel([0.146733, -0.792929, -2.792159, -1.127301, 1.570796, 1.717529],accel_mss,speed_ms,0,blend_radius_m)
  movel([0.142223, -0.794583, -2.791882, -1.125924, 1.570796, 1.713020],accel_mss,speed_ms,0,blend_radius_m)
  movel([0.142758, -0.796773, -2.791513, -1.124103, 1.570796, 1.713554],accel_mss,speed_ms,0,blend_radius_m)
  movel([0.143619, -0.799117, -2.791116, -1.122156, 1.570796, 1.714415],accel_mss,speed_ms,0,blend_radius_m)
  movel([0.144902, -0.801444, -2.790719, -1.120226, 1.570796, 1.715698],accel_mss,speed_ms,0,blend_radius_m)
  movel([0.146705, -0.803590, -2.790350, -1.118450, 1.570796, 1.717501],accel_mss,speed_ms,0,blend_radius_m)
  movel([0.152042, -0.805679, -2.789988, -1.116722, 1.570796, 1.722838],accel_mss,speed_ms,0,blend_radius_m)
  movel([0.154980, -0.807003, -2.789758, -1.115628, 1.570796, 1.725776],accel_mss,speed_ms,0,blend_radius_m)
  movel([0.155811, -0.807709, -2.789635, -1.115046, 1.570796, 1.726607],accel_mss,speed_ms,0,blend_radius_m)
  movel([0.155954, -0.808432, -2.789508, -1.114449, 1.570796, 1.726751],accel_mss,speed_ms,0,blend_radius_m)
  movel([0.155514, -0.809285, -2.789359, -1.113746, 1.570796, 1.726310],accel_mss,speed_ms,0,blend_radius_m)
  movel([0.154880, -0.810099, -2.789215, -1.113074, 1.570796, 1.725676],accel_mss,speed_ms,0,blend_radius_m)
  movel([0.153372, -0.811356, -2.788994, -1.112039, 1.570796, 1.724168],accel_mss,speed_ms,0,blend_radius_m)
  movel([0.152148, -0.811911, -2.788896, -1.111582, 1.570796, 1.722944],accel_mss,speed_ms,0,blend_radius_m)
  movel([0.150940, -0.812222, -2.788841, -1.111326, 1.570796, 1.721736],accel_mss,speed_ms,0,blend_radius_m)
  movel([0.148664, -0.812617, -2.788771, -1.111001, 1.570796, 1.719461],accel_mss,speed_ms,0,blend_radius_m)
  movel([0.149487, -0.815555, -2.788248, -1.108586, 1.570796, 1.720283],accel_mss,speed_ms,0,blend_radius_m)
  movel([0.150580, -0.818226, -2.787768, -1.106395, 1.570796, 1.721377],accel_mss,speed_ms,0,blend_radius_m)
  movel([0.151941, -0.820619, -2.787335, -1.104435, 1.570796, 1.722738],accel_mss,speed_ms,0,blend_radius_m)
  movel([0.153547, -0.822737, -2.786949, -1.102703, 1.570796, 1.724344],accel_mss,speed_ms,0,blend_radius_m)
  movel([0.155518, -0.824369, -2.786650, -1.101370, 1.570796, 1.726315],accel_mss,speed_ms,0,blend_radius_m)
  movel([0.157892, -0.825466, -2.786448, -1.100475, 1.570796, 1.728688],accel_mss,speed_ms,0,blend_radius_m)
  movel([0.163164, -0.826884, -2.786186, -1.099318, 1.570796, 1.733961],accel_mss,speed_ms,0,blend_radius_m)
  movel([0.164477, -0.827614, -2.786051, -1.098723, 1.570796, 1.735273],accel_mss,speed_ms,0,blend_radius_m)
  movel([0.164731, -0.828352, -2.785915, -1.098123, 1.570796, 1.735527],accel_mss,speed_ms,0,blend_radius_m)
  movel([0.164486, -0.829419, -2.785716, -1.097254, 1.570796, 1.735282],accel_mss,speed_ms,0,blend_radius_m)
  movel([0.163859, -0.830453, -2.785523, -1.096413, 1.570796, 1.734656],accel_mss,speed_ms,0,blend_radius_m)
  movel([0.163012, -0.831369, -2.785351, -1.095669, 1.570796, 1.733808],accel_mss,speed_ms,0,blend_radius_m)
  movel([0.161071, -0.832811, -2.785080, -1.094498, 1.570796, 1.731867],accel_mss,speed_ms,0,blend_radius_m)
  movel([0.158538, -0.834202, -2.784818, -1.093369, 1.570796, 1.729334],accel_mss,speed_ms,0,blend_radius_m)
  movel([0.156117, -0.835242, -2.784621, -1.092526, 1.570796, 1.726913],accel_mss,speed_ms,0,blend_radius_m)
  movel([0.153793, -0.835986, -2.784480, -1.091923, 1.570796, 1.724589],accel_mss,speed_ms,0,blend_radius_m)
  movel([0.151559, -0.836468, -2.784388, -1.091533, 1.570796, 1.722355],accel_mss,speed_ms,0,blend_radius_m)
  movel([0.152827, -0.838488, -2.784003, -1.089899, 1.570796, 1.723624],accel_mss,speed_ms,0,blend_radius_m)
  movel([0.154404, -0.840131, -2.783688, -1.088571, 1.570796, 1.725200],accel_mss,speed_ms,0,blend_radius_m)
  movel([0.156283, -0.841354, -2.783452, -1.087583, 1.570796, 1.727080],accel_mss,speed_ms,0,blend_radius_m)
  movel([0.158458, -0.842122, -2.783303, -1.086963, 1.570796, 1.729255],accel_mss,speed_ms,0,blend_radius_m)
  movel([0.160934, -0.842390, -2.783252, -1.086748, 1.570796, 1.731730],accel_mss,speed_ms,0,blend_radius_m)
  movel([0.163710, -0.842116, -2.783305, -1.086968, 1.570796, 1.734507],accel_mss,speed_ms,0,blend_radius_m)
  movel([0.166787, -0.841254, -2.783471, -1.087664, 1.570796, 1.737583],accel_mss,speed_ms,0,blend_radius_m)
  movel([0.170171, -0.839761, -2.783759, -1.088870, 1.570796, 1.740967],accel_mss,speed_ms,0,blend_radius_m)
  speed_ms = 0.005
  movel([0.170171, -0.831312, -2.777505, -1.103572, 1.570796, 1.740967],accel_mss,speed_ms,0,blend_radius_m)
  speed_ms = 0.040
  movel([0.185325, -0.808402, -2.781729, -1.122258, 1.570796, 1.756121],accel_mss,speed_ms,0,blend_radius_m)
  speed_ms = 0.005
  movel([0.185325, -0.816634, -2.788054, -1.107701, 1.570796, 1.756121],accel_mss,speed_ms,0,blend_radius_m)
  speed_ms = 0.025
  movel([0.179130, -0.816481, -2.788082, -1.107826, 1.570796, 1.749926],accel_mss,speed_ms,0,blend_radius_m)
  movel([0.176504, -0.816112, -2.788148, -1.108129, 1.570796, 1.747300],accel_mss,speed_ms,0,blend_radius_m)
  movel([0.174175, -0.815445, -2.788267, -1.108676, 1.570796, 1.744971],accel_mss,speed_ms,0,blend_radius_m)
  movel([0.172123, -0.814400, -2.788454, -1.109535, 1.570796, 1.742919],accel_mss,speed_ms,0,blend_radius_m)
  movel([0.170335, -0.812901, -2.788720, -1.110768, 1.570796, 1.741131],accel_mss,speed_ms,0,blend_radius_m)
  movel([0.168788, -0.810874, -2.789079, -1.112436, 1.570796, 1.739584],accel_mss,speed_ms,0,blend_radius_m)
  movel([0.167475, -0.808237, -2.789542, -1.114610, 1.570796, 1.738271],accel_mss,speed_ms,0,blend_radius_m)
  movel([0.165467, -0.802003, -2.790623, -1.119764, 1.570796, 1.736263],accel_mss,speed_ms,0,blend_radius_m)
  movel([0.164156, -0.795093, -2.791797, -1.125500, 1.570796, 1.734952],accel_mss,speed_ms,0,blend_radius_m)
  movel([0.163481, -0.787589, -2.793043, -1.131756, 1.570796, 1.734277],accel_mss,speed_ms,0,blend_radius_m)
  movel([0.163370, -0.779597, -2.794339, -1.138452, 1.570796, 1.734166],accel_mss,speed_ms,0,blend_radius_m)
  movel([0.163693, -0.772714, -2.795430, -1.144245, 1.570796, 1.734489],accel_mss,speed_ms,0,blend_radius_m)
  movel([0.164351, -0.765561, -2.796538, -1.150290, 1.570796, 1.735147],accel_mss,speed_ms,0,blend_radius_m)
  movel([0.166427, -0.750590, -2.798776, -1.163023, 1.570796, 1.737223],accel_mss,speed_ms,0,blend_radius_m)
  movel([0.175526, -0.696644, -2.805963, -1.209781, 1.570796, 1.746322],accel_mss,speed_ms,0,blend_radius_m)
  movel([0.177448, -0.685048, -2.807336, -1.220005, 1.570796, 1.748244],accel_mss,speed_ms,0,blend_radius_m)
  movel([0.179180, -0.673475, -2.808648, -1.230267, 1.570796, 1.749976],accel_mss,speed_ms,0,blend_radius_m)
  movel([0.180554, -0.662095, -2.809881, -1.240412, 1.570796, 1.751350],accel_mss,speed_ms,0,blend_radius_m)
  movel([0.181390, -0.651075, -2.811024, -1.250291, 1.570796, 1.752186],accel_mss,speed_ms,0,blend_radius_m)
  movel([0.181508, -0.640597, -2.812063, -1.259730, 1.570796, 1.752305],accel_mss,speed_ms,0,blend_radius_m)
  movel([0.180716, -0.630855, -2.812989, -1.268545, 1.570796, 1.751512],accel_mss,speed_ms,0,blend_radius_m)
  movel([0.179492, -0.624313, -2.813589, -1.274488, 1.570796, 1.750288],accel_mss,speed_ms,0,blend_radius_m)
  movel([0.177674, -0.618108, -2.814142, -1.280139, 1.570796, 1.748470],accel_mss,speed_ms,0,blend_radius_m)
  movel([0.175212, -0.612418, -2.814635, -1.285336, 1.570796, 1.746008],accel_mss,speed_ms,0,blend_radius_m)
  movel([0.172054, -0.607420, -2.815058, -1.289910, 1.570796, 1.742851],accel_mss,speed_ms,0,blend_radius_m)
  movel([0.168163, -0.603283, -2.815401, -1.293705, 1.570796, 1.738959],accel_mss,speed_ms,0,blend_radius_m)
  movel([0.163499, -0.600172, -2.815654, -1.296562, 1.570796, 1.734295],accel_mss,speed_ms,0,blend_radius_m)
  movel([0.158021, -0.598271, -2.815807, -1.298310, 1.570796, 1.728817],accel_mss,speed_ms,0,blend_radius_m)
  movel([0.151716, -0.597732, -2.815851, -1.298807, 1.570796, 1.722513],accel_mss,speed_ms,0,blend_radius_m)
  movel([0.148431, -0.598051, -2.815825, -1.298513, 1.570796, 1.719227],accel_mss,speed_ms,0,blend_radius_m)
  movel([0.144882, -0.598822, -2.815763, -1.297803, 1.570796, 1.715678],accel_mss,speed_ms,0,blend_radius_m)
  movel([0.141095, -0.600068, -2.815663, -1.296658, 1.570796, 1.711892],accel_mss,speed_ms,0,blend_radius_m)
  movel([0.137112, -0.601797, -2.815523, -1.295069, 1.570796, 1.707908],accel_mss,speed_ms,0,blend_radius_m)
  movel([0.132975, -0.604009, -2.815342, -1.293039, 1.570796, 1.703772],accel_mss,speed_ms,0,blend_radius_m)
  movel([0.128708, -0.606727, -2.815116, -1.290545, 1.570796, 1.699505],accel_mss,speed_ms,0,blend_radius_m)
  movel([0.124362, -0.609943, -2.814846, -1.287599, 1.570796, 1.695159],accel_mss,speed_ms,0,blend_radius_m)
  movel([0.119974, -0.613671, -2.814528, -1.284190, 1.570796, 1.690770],accel_mss,speed_ms,0,blend_radius_m)
  speed_ms = 0.005
  movel([0.119974, -0.608102, -2.807721, -1.296566, 1.570796, 1.690770],accel_mss,speed_ms,0,blend_radius_m)
  speed_ms = 0.040
  movel([0.105668, -0.595567, -2.808765, -1.308057, 1.570796, 1.676464],accel_mss,speed_ms,0,blend_radius_m)
  speed_ms = 0.005
  movel([0.105668, -0.600928, -2.815593, -1.295868, 1.570796, 1.676464],accel_mss,speed_ms,0,blend_radius_m)
  speed_ms = 0.025
  movel([0.105208, -0.598577, -2.815783, -1.298029, 1.570796, 1.676004],accel_mss,speed_ms,0,blend_radius_m)
  movel([0.105101, -0.595921, -2.815994, -1.300473, 1.570796, 1.675897],accel_mss,speed_ms,0,blend_radius_m)
  movel([0.105749, -0.589893, -2.816465, -1.306031, 1.570796, 1.676545],accel_mss,speed_ms,0,blend_radius_m)
  movel([0.107230, -0.583192, -2.816971, -1.312227, 1.570796, 1.678026],accel_mss,speed_ms,0,blend_radius_m)
  movel([0.109136, -0.576203, -2.817480, -1.318706, 1.570796, 1.679932],accel_mss,speed_ms,0,blend_radius_m)
  speed_ms = 0.005
  movel([0.109136, -0.571256, -2.810615, -1.330518, 1.570796, 1.679932],accel_mss,speed_ms,0,blend_radius_m)
  speed_ms = 0.040
  movel([0.118580, -0.567918, -2.810851, -1.333621, 1.570796, 1.689376],accel_mss,speed_ms,0,blend_radius_m)
  speed_ms = 0.005
  movel([0.118580, -0.572806, -2.817721, -1.321862, 1.570796, 1.689376],accel_mss,speed_ms,0,blend_radius_m)
  speed_ms = 0.025
  movel([0.117402, -0.571397, -2.817820, -1.323172, 1.570796, 1.688198],accel_mss,speed_ms,0,blend_radius_m)
  movel([0.116582, -0.569671, -2.817939, -1.324778, 1.570796, 1.687379],accel_mss,speed_ms,0,blend_radius_m)
  movel([0.115918, -0.565351, -2.818234, -1.328804, 1.570796, 1.686715],accel_mss,speed_ms,0,blend_radius_m)
  movel([0.116427, -0.560033, -2.818587, -1.333768, 1.570796, 1.687223],accel_mss,speed_ms,0,blend_radius_m)
  movel([0.117944, -0.553895, -2.818982, -1.339512, 1.570796, 1.688741],accel_mss,speed_ms,0,blend_radius_m)
  movel([0.120304, -0.547129, -2.819401, -1.345859, 1.570796, 1.691100],accel_mss,speed_ms,0,blend_radius_m)
  movel([0.123332, -0.539934, -2.819828, -1.352628, 1.570796, 1.694129],accel_mss,speed_ms,0,blend_radius_m)
  movel([0.126853, -0.532508, -2.820248, -1.359633, 1.570796, 1.697649],accel_mss,speed_ms,0,blend_radius_m)
  movel([0.130680, -0.525067, -2.820649, -1.366673, 1.570796, 1.701476],accel_mss,speed_ms,0,blend_radius_m)
  speed_ms = 0.005
  movel([0.130680, -0.521025, -2.813720, -1.377644, 1.570796, 1.701476],accel_mss,speed_ms,0,blend_radius_m)
  speed_ms = 0.040
  movel([0.181260, -0.451275, -2.816496, -1.444618, 1.570796, 1.752057],accel_mss,speed_ms,0,blend_radius_m)
  speed_ms = 0.005
  movel([0.181260, -0.453974, -2.823484, -1.434931, 1.570796, 1.752057],accel_mss,speed_ms,0,blend_radius_m)
  speed_ms = 0.025
  movel([0.176078, -0.459840, -2.823317, -1.429232, 1.570796, 1.746874],accel_mss,speed_ms,0,blend_radius_m)
  movel([0.170926, -0.466016, -2.823129, -1.423245, 1.570796, 1.741722],accel_mss,speed_ms,0,blend_radius_m)
  movel([0.165890, -0.472402, -2.822920, -1.417067, 1.570796, 1.736686],accel_mss,speed_ms,0,blend_radius_m)
  movel([0.161028, -0.478924, -2.822692, -1.410773, 1.570796, 1.731824],accel_mss,speed_ms,0,blend_radius_m)
  movel([0.156423, -0.485495, -2.822447, -1.404447, 1.570796, 1.727219],accel_mss,speed_ms,0,blend_radius_m)
  movel([0.152136, -0.492027, -2.822189, -1.398173, 1.570796, 1.722932],accel_mss,speed_ms,0,blend_radius_m)
  movel([0.148234, -0.498450, -2.821920, -1.392019, 1.570796, 1.719030],accel_mss,speed_ms,0,blend_radius_m)
  movel([0.144778, -0.504688, -2.821645, -1.386056, 1.570796, 1.715575],accel_mss,speed_ms,0,blend_radius_m)
  movel([0.141828, -0.510657, -2.821369, -1.380363, 1.570796, 1.712624],accel_mss,speed_ms,0,blend_radius_m)
  movel([0.139435, -0.516300, -2.821096, -1.374994, 1.570796, 1.710232],accel_mss,speed_ms,0,blend_radius_m)
  movel([0.137657, -0.521542, -2.820832, -1.370015, 1.570796, 1.708453],accel_mss,speed_ms,0,blend_radius_m)
  movel([0.136544, -0.526318, -2.820583, -1.365488, 1.570796, 1.707340],accel_mss,speed_ms,0,blend_radius_m)
  movel([0.136155, -0.530558, -2.820355, -1.361476, 1.570796, 1.706952],accel_mss,speed_ms,0,blend_radius_m)
  movel([0.136543, -0.534201, -2.820154, -1.358034, 1.570796, 1.707339],accel_mss,speed_ms,0,blend_radius_m)
  movel([0.137752, -0.537189, -2.819985, -1.355215, 1.570796, 1.708548],accel_mss,speed_ms,0,blend_radius_m)
  movel([0.139843, -0.539457, -2.819855, -1.353077, 1.570796, 1.710639],accel_mss,speed_ms,0,blend_radius_m)
  speed_ms = 0.005
  movel([0.139843, -0.535154, -2.812942, -1.364293, 1.570796, 1.710639],accel_mss,speed_ms,0,blend_radius_m)
  speed_ms = 0.040
  movel([0.162855, -0.510032, -2.814274, -1.388084, 1.570796, 1.733652],accel_mss,speed_ms,0,blend_radius_m)
  speed_ms = 0.005
  movel([0.162855, -0.513869, -2.821215, -1.377306, 1.570796, 1.733652],accel_mss,speed_ms,0,blend_radius_m)
  speed_ms = 0.025
  movel([0.162384, -0.510995, -2.821353, -1.380041, 1.570796, 1.733180],accel_mss,speed_ms,0,blend_radius_m)
  movel([0.162288, -0.507765, -2.821504, -1.383120, 1.570796, 1.733084],accel_mss,speed_ms,0,blend_radius_m)
  movel([0.162565, -0.504214, -2.821666, -1.386509, 1.570796, 1.733362],accel_mss,speed_ms,0,blend_radius_m)
  movel([0.163216, -0.500361, -2.821837, -1.390191, 1.570796, 1.734012],accel_mss,speed_ms,0,blend_radius_m)
  movel([0.164233, -0.496243, -2.822014, -1.394132, 1.570796, 1.735029],accel_mss,speed_ms,0,blend_radius_m)
  movel([0.165623, -0.491879, -2.822195, -1.398315, 1.570796, 1.736419],accel_mss,speed_ms,0,blend_radius_m)
  movel([0.167387, -0.487288, -2.822378, -1.402723, 1.570796, 1.738183],accel_mss,speed_ms,0,blend_radius_m)
  movel([0.169516, -0.482514, -2.822560, -1.407315, 1.570796, 1.740313],accel_mss,speed_ms,0,blend_radius_m)
  movel([0.172012, -0.477577, -2.822740, -1.412072, 1.570796, 1.742809],accel_mss,speed_ms,0,blend_radius_m)
  movel([0.174881, -0.472499, -2.822916, -1.416973, 1.570796, 1.745678],accel_mss,speed_ms,0,blend_radius_m)
  movel([0.178106, -0.467332, -2.823087, -1.421970, 1.570796, 1.748902],accel_mss,speed_ms,0,blend_radius_m)
  movel([0.181701, -0.462081, -2.823250, -1.427058, 1.570796, 1.752497],accel_mss,speed_ms,0,blend_radius_m)
  movel([0.185655, -0.456788, -2.823405, -1.432195, 1.570796, 1.756451],accel_mss,speed_ms,0,blend_radius_m)
  movel([0.189965, -0.451486, -2.823551, -1.437352, 1.570796, 1.760761],accel_mss,speed_ms,0,blend_radius_m)
  movel([0.194624, -0.446213, -2.823686, -1.442490, 1.570796, 1.765421],accel_mss,speed_ms,0,blend_radius_m)
  movel([0.199621, -0.441004, -2.823810, -1.447575, 1.570796, 1.770417],accel_mss,speed_ms,0,blend_radius_m)
  movel([0.204634, -0.436212, -2.823916, -1.452261, 1.570796, 1.775430],accel_mss,speed_ms,0,blend_radius_m)
  movel([0.209620, -0.431863, -2.824006, -1.456520, 1.570796, 1.780416],accel_mss,speed_ms,0,blend_radius_m)
  movel([0.214539, -0.427961, -2.824081, -1.460347, 1.570796, 1.785336],accel_mss,speed_ms,0,blend_radius_m)
  movel([0.219373, -0.424507, -2.824142, -1.463739, 1.570796, 1.790170],accel_mss,speed_ms,0,blend_radius_m)
  movel([0.224084, -0.421505, -2.824193, -1.466691, 1.570796, 1.794880],accel_mss,speed_ms,0,blend_radius_m)
  movel([0.228628, -0.418970, -2.824233, -1.469186, 1.570796, 1.799425],accel_mss,speed_ms,0,blend_radius_m)
  movel([0.232995, -0.416879, -2.824265, -1.471245, 1.570796, 1.803792],accel_mss,speed_ms,0,blend_radius_m)
  movel([0.237129, -0.415258, -2.824288, -1.472843, 1.570796, 1.807925],accel_mss,speed_ms,0,blend_radius_m)
  movel([0.241016, -0.414095, -2.824304, -1.473990, 1.570796, 1.811812],accel_mss,speed_ms,0,blend_radius_m)
  movel([0.247935, -0.413121, -2.824318, -1.474951, 1.570796, 1.818732],accel_mss,speed_ms,0,blend_radius_m)
  movel([0.250900, -0.413314, -2.824315, -1.474760, 1.570796, 1.821697],accel_mss,speed_ms,0,blend_radius_m)
  movel([0.255753, -0.415004, -2.824292, -1.473093, 1.570796, 1.826549],accel_mss,speed_ms,0,blend_radius_m)
  movel([0.257590, -0.416485, -2.824270, -1.471633, 1.570796, 1.828387],accel_mss,speed_ms,0,blend_radius_m)
  movel([0.259001, -0.418384, -2.824242, -1.469763, 1.570796, 1.829798],accel_mss,speed_ms,0,blend_radius_m)
  speed_ms = 0.005
  movel([0.259001, -0.416389, -2.817239, -1.478762, 1.570796, 1.829798],accel_mss,speed_ms,0,blend_radius_m)
  speed_ms = 0.040
  movel([0.274724, -0.429162, -2.817016, -1.466211, 1.570796, 1.845520],accel_mss,speed_ms,0,blend_radius_m)
  speed_ms = 0.005
  movel([0.274724, -0.431417, -2.824015, -1.456957, 1.570796, 1.845520],accel_mss,speed_ms,0,blend_radius_m)
  speed_ms = 0.025
  movel([0.272812, -0.428276, -2.824075, -1.460038, 1.570796, 1.843609],accel_mss,speed_ms,0,blend_radius_m)
  movel([0.269936, -0.426281, -2.824111, -1.461997, 1.570796, 1.840732],accel_mss,speed_ms,0,blend_radius_m)
  movel([0.266170, -0.425428, -2.824126, -1.462835, 1.570796, 1.836967],accel_mss,speed_ms,0,blend_radius_m)
  movel([0.261578, -0.425716, -2.824121, -1.462552, 1.570796, 1.832374],accel_mss,speed_ms,0,blend_radius_m)
  movel([0.256264, -0.427118, -2.824096, -1.461175, 1.570796, 1.827060],accel_mss,speed_ms,0,blend_radius_m)
  movel([0.250302, -0.429626, -2.824049, -1.458714, 1.570796, 1.821099],accel_mss,speed_ms,0,blend_radius_m)
  movel([0.243802, -0.433205, -2.823979, -1.455205, 1.570796, 1.814599],accel_mss,speed_ms,0,blend_radius_m)
  movel([0.236850, -0.437832, -2.823881, -1.450676, 1.570796, 1.807647],accel_mss,speed_ms,0,blend_radius_m)
  movel([0.229570, -0.443455, -2.823753, -1.445181, 1.570796, 1.800366],accel_mss,speed_ms,0,blend_radius_m)
  movel([0.222137, -0.449962, -2.823591, -1.438836, 1.570796, 1.792933],accel_mss,speed_ms,0,blend_radius_m)
  movel([0.214847, -0.457117, -2.823396, -1.431876, 1.570796, 1.785644],accel_mss,speed_ms,0,blend_radius_m)
  movel([0.208004, -0.464688, -2.823170, -1.424530, 1.570796, 1.778801],accel_mss,speed_ms,0,blend_radius_m)
  movel([0.201871, -0.472470, -2.822917, -1.417002, 1.570796, 1.772667],accel_mss,speed_ms,0,blend_radius_m)
  movel([0.199162, -0.476367, -2.822783, -1.413239, 1.570796, 1.769958],accel_mss,speed_ms,0,blend_radius_m)
  movel([0.196726, -0.480235, -2.822644, -1.409509, 1.570796, 1.767523],accel_mss,speed_ms,0,blend_radius_m)
  movel([0.194595, -0.484056, -2.822502, -1.405831, 1.570796, 1.765391],accel_mss,speed_ms,0,blend_radius_m)
  movel([0.192805, -0.487805, -2.822357, -1.402226, 1.570796, 1.763601],accel_mss,speed_ms,0,blend_radius_m)
  movel([0.191376, -0.491457, -2.822212, -1.398720, 1.570796, 1.762173],accel_mss,speed_ms,0,blend_radius_m)
  movel([0.190353, -0.494977, -2.822067, -1.395345, 1.570796, 1.761149],accel_mss,speed_ms,0,blend_radius_m)
  speed_ms = 0.005
  movel([0.190353, -0.491492, -2.815109, -1.405788, 1.570796, 1.761149],accel_mss,speed_ms,0,blend_radius_m)
  speed_ms = 0.040
  movel([0.225557, -0.480547, -2.815543, -1.416299, 1.570796, 1.796354],accel_mss,speed_ms,0,blend_radius_m)
  speed_ms = 0.005
  movel([0.225557, -0.483821, -2.822511, -1.406057, 1.570796, 1.796354],accel_mss,speed_ms,0,blend_radius_m)
  speed_ms = 0.025
  movel([0.230532, -0.478358, -2.822712, -1.411318, 1.570796, 1.801329],accel_mss,speed_ms,0,blend_radius_m)
  movel([0.235675, -0.473359, -2.822887, -1.416143, 1.570796, 1.806472],accel_mss,speed_ms,0,blend_radius_m)
  movel([0.240904, -0.468850, -2.823038, -1.420501, 1.570796, 1.811700],accel_mss,speed_ms,0,blend_radius_m)
  movel([0.246113, -0.464881, -2.823164, -1.424344, 1.570796, 1.816909],accel_mss,speed_ms,0,blend_radius_m)
  movel([0.251210, -0.461482, -2.823268, -1.427639, 1.570796, 1.822007],accel_mss,speed_ms,0,blend_radius_m)
  movel([0.256093, -0.458688, -2.823351, -1.430351, 1.570796, 1.826889],accel_mss,speed_ms,0,blend_radius_m)
  movel([0.260676, -0.456527, -2.823413, -1.432449, 1.570796, 1.831472],accel_mss,speed_ms,0,blend_radius_m)
  movel([0.264851, -0.455034, -2.823455, -1.433900, 1.570796, 1.835647],accel_mss,speed_ms,0,blend_radius_m)
  movel([0.269216, -0.454288, -2.823475, -1.434626, 1.570796, 1.840012],accel_mss,speed_ms,0,blend_radius_m)
  movel([0.272323, -0.454879, -2.823459, -1.434051, 1.570796, 1.843120],accel_mss,speed_ms,0,blend_radius_m)
  movel([0.274310, -0.456660, -2.823409, -1.432320, 1.570796, 1.845106],accel_mss,speed_ms,0,blend_radius_m)
  movel([0.275291, -0.459498, -2.823327, -1.429564, 1.570796, 1.846087],accel_mss,speed_ms,0,blend_radius_m)
  movel([0.275404, -0.463233, -2.823215, -1.425941, 1.570796, 1.846201],accel_mss,speed_ms,0,blend_radius_m)
  movel([0.274782, -0.467729, -2.823074, -1.421586, 1.570796, 1.845579],accel_mss,speed_ms,0,blend_radius_m)
  movel([0.273555, -0.472838, -2.822905, -1.416646, 1.570796, 1.844351],accel_mss,speed_ms,0,blend_radius_m)
  movel([0.271863, -0.478411, -2.822710, -1.411268, 1.570796, 1.842660],accel_mss,speed_ms,0,blend_radius_m)
  speed_ms = 0.005
  movel([0.271863, -0.475240, -2.815739, -1.421411, 1.570796, 1.842660],accel_mss,speed_ms,0,blend_radius_m)
  speed_ms = 0.040
  movel([0.237934, -0.495293, -2.814948, -1.402148, 1.570796, 1.808730],accel_mss,speed_ms,0,blend_radius_m)
  speed_ms = 0.005
  movel([0.237934, -0.498851, -2.821903, -1.391636, 1.570796, 1.808730],accel_mss,speed_ms,0,blend_radius_m)
  speed_ms = 0.025
  movel([0.242451, -0.496479, -2.822004, -1.393906, 1.570796, 1.813247],accel_mss,speed_ms,0,blend_radius_m)
  movel([0.246530, -0.494816, -2.822074, -1.395500, 1.570796, 1.817326],accel_mss,speed_ms,0,blend_radius_m)
  movel([0.250167, -0.493844, -2.822114, -1.396431, 1.570796, 1.820964],accel_mss,speed_ms,0,blend_radius_m)
  movel([0.253371, -0.493515, -2.822128, -1.396746, 1.570796, 1.824168],accel_mss,speed_ms,0,blend_radius_m)
  movel([0.256145, -0.493804, -2.822116, -1.396469, 1.570796, 1.826941],accel_mss,speed_ms,0,blend_radius_m)
  movel([0.258492, -0.494668, -2.822080, -1.395641, 1.570796, 1.829288],accel_mss,speed_ms,0,blend_radius_m)
  movel([0.260428, -0.496068, -2.822021, -1.394300, 1.570796, 1.831224],accel_mss,speed_ms,0,blend_radius_m)
  movel([0.261949, -0.497976, -2.821940, -1.392473, 1.570796, 1.832745],accel_mss,speed_ms,0,blend_radius_m)
  movel([0.263082, -0.500341, -2.821838, -1.390210, 1.570796, 1.833878],accel_mss,speed_ms,0,blend_radius_m)
  movel([0.263834, -0.503122, -2.821715, -1.387552, 1.570796, 1.834630],accel_mss,speed_ms,0,blend_radius_m)
  movel([0.264212, -0.506287, -2.821572, -1.384530, 1.570796, 1.835008],accel_mss,speed_ms,0,blend_radius_m)
  movel([0.264237, -0.509786, -2.821410, -1.381194, 1.570796, 1.835033],accel_mss,speed_ms,0,blend_radius_m)
  movel([0.263917, -0.513585, -2.821228, -1.377575, 1.570796, 1.834713],accel_mss,speed_ms,0,blend_radius_m)
  movel([0.262305, -0.521909, -2.820813, -1.369667, 1.570796, 1.833101],accel_mss,speed_ms,0,blend_radius_m)
  movel([0.261033, -0.526363, -2.820581, -1.365445, 1.570796, 1.831830],accel_mss,speed_ms,0,blend_radius_m)
  movel([0.260911, -0.525245, -2.820640, -1.366504, 1.570796, 1.831708],accel_mss,speed_ms,0,blend_radius_m)
  speed_ms = 0.005
  movel([0.260911, -0.521200, -2.813710, -1.377479, 1.570796, 1.831708],accel_mss,speed_ms,0,blend_radius_m)
  speed_ms = 0.040
  movel([0.286425, -0.519761, -2.813786, -1.378843, 1.570796, 1.857221],accel_mss,speed_ms,0,blend_radius_m)
  speed_ms = 0.005
  movel([0.286425, -0.523780, -2.820716, -1.367893, 1.570796, 1.857221],accel_mss,speed_ms,0,blend_radius_m)
  speed_ms = 0.025
  movel([0.281721, -0.531053, -2.820328, -1.361008, 1.570796, 1.852517],accel_mss,speed_ms,0,blend_radius_m)
  movel([0.277579, -0.538222, -2.819926, -1.354241, 1.570796, 1.848375],accel_mss,speed_ms,0,blend_radius_m)
  movel([0.273882, -0.545266, -2.819513, -1.347610, 1.570796, 1.844679],accel_mss,speed_ms,0,blend_radius_m)
  movel([0.270506, -0.552173, -2.819090, -1.341126, 1.570796, 1.841302],accel_mss,speed_ms,0,blend_radius_m)
  movel([0.267119, -0.559621, -2.818614, -1.334154, 1.570796, 1.837915],accel_mss,speed_ms,0,blend_radius_m)
  movel([0.265729, -0.563180, -2.818380, -1.330829, 1.570796, 1.836525],accel_mss,speed_ms,0,blend_radius_m)
  movel([0.264664, -0.566551, -2.818153, -1.327685, 1.570796, 1.835460],accel_mss,speed_ms,0,blend_radius_m)
  movel([0.264005, -0.569666, -2.817940, -1.324783, 1.570796, 1.834801],accel_mss,speed_ms,0,blend_radius_m)
  movel([0.263849, -0.572391, -2.817750, -1.322248, 1.570796, 1.834645],accel_mss,speed_ms,0,blend_radius_m)
  movel([0.264284, -0.574553, -2.817598, -1.320239, 1.570796, 1.835080],accel_mss,speed_ms,0,blend_radius_m)
  movel([0.265378, -0.576013, -2.817494, -1.318883, 1.570796, 1.836174],accel_mss,speed_ms,0,blend_radius_m)
  movel([0.268144, -0.577019, -2.817422, -1.317948, 1.570796, 1.838940],accel_mss,speed_ms,0,blend_radius_m)
  movel([0.269503, -0.577541, -2.817384, -1.317464, 1.570796, 1.840299],accel_mss,speed_ms,0,blend_radius_m)
  movel([0.270510, -0.578493, -2.817315, -1.316581, 1.570796, 1.841306],accel_mss,speed_ms,0,blend_radius_m)
  movel([0.270926, -0.580427, -2.817174, -1.314788, 1.570796, 1.841723],accel_mss,speed_ms,0,blend_radius_m)
  movel([0.270622, -0.583206, -2.816970, -1.312213, 1.570796, 1.841419],accel_mss,speed_ms,0,blend_radius_m)
  movel([0.269763, -0.586603, -2.816715, -1.309070, 1.570796, 1.840560],accel_mss,speed_ms,0,blend_radius_m)
  movel([0.268504, -0.590388, -2.816427, -1.305575, 1.570796, 1.839300],accel_mss,speed_ms,0,blend_radius_m)
  movel([0.265395, -0.598243, -2.815810, -1.298336, 1.570796, 1.836191],accel_mss,speed_ms,0,blend_radius_m)
  movel([0.255783, -0.620300, -2.813948, -1.278141, 1.570796, 1.826579],accel_mss,speed_ms,0,blend_radius_m)
  movel([0.249309, -0.635304, -2.812571, -1.264514, 1.570796, 1.820106],accel_mss,speed_ms,0,blend_radius_m)
  movel([0.247618, -0.639771, -2.812143, -1.260475, 1.570796, 1.818415],accel_mss,speed_ms,0,blend_radius_m)
  movel([0.246095, -0.644412, -2.811690, -1.256287, 1.570796, 1.816891],accel_mss,speed_ms,0,blend_radius_m)
  movel([0.243703, -0.653805, -2.810745, -1.247839, 1.570796, 1.814500],accel_mss,speed_ms,0,blend_radius_m)
  movel([0.242917, -0.658353, -2.810275, -1.243761, 1.570796, 1.813713],accel_mss,speed_ms,0,blend_radius_m)
  movel([0.242456, -0.662667, -2.809821, -1.239901, 1.570796, 1.813252],accel_mss,speed_ms,0,blend_radius_m)
  movel([0.242353, -0.666651, -2.809394, -1.236344, 1.570796, 1.813149],accel_mss,speed_ms,0,blend_radius_m)
  movel([0.242645, -0.670213, -2.809007, -1.233169, 1.570796, 1.813442],accel_mss,speed_ms,0,blend_radius_m)
  movel([0.243374, -0.673244, -2.808673, -1.230471, 1.570796, 1.814170],accel_mss,speed_ms,0,blend_radius_m)
  movel([0.244568, -0.675669, -2.808404, -1.228317, 1.570796, 1.815364],accel_mss,speed_ms,0,blend_radius_m)
  movel([0.246276, -0.677375, -2.808212, -1.226802, 1.570796, 1.817072],accel_mss,speed_ms,0,blend_radius_m)
  movel([0.248533, -0.678274, -2.808111, -1.226004, 1.570796, 1.819329],accel_mss,speed_ms,0,blend_radius_m)
  movel([0.251378, -0.678269, -2.808111, -1.226008, 1.570796, 1.822174],accel_mss,speed_ms,0,blend_radius_m)
  movel([0.254864, -0.677254, -2.808226, -1.226909, 1.570796, 1.825661],accel_mss,speed_ms,0,blend_radius_m)
  movel([0.259038, -0.675131, -2.808464, -1.228794, 1.570796, 1.829835],accel_mss,speed_ms,0,blend_radius_m)
  movel([0.263958, -0.671786, -2.808834, -1.231768, 1.570796, 1.834754],accel_mss,speed_ms,0,blend_radius_m)
  movel([0.267886, -0.668616, -2.809181, -1.234592, 1.570796, 1.838682],accel_mss,speed_ms,0,blend_radius_m)
  movel([0.271783, -0.665089, -2.809562, -1.237738, 1.570796, 1.842579],accel_mss,speed_ms,0,blend_radius_m)
  movel([0.275661, -0.661254, -2.809970, -1.241165, 1.570796, 1.846457],accel_mss,speed_ms,0,blend_radius_m)
  movel([0.279521, -0.657170, -2.810398, -1.244821, 1.570796, 1.850318],accel_mss,speed_ms,0,blend_radius_m)
  movel([0.287206, -0.648497, -2.811284, -1.252609, 1.570796, 1.858002],accel_mss,speed_ms,0,blend_radius_m)
  movel([0.294865, -0.639552, -2.812164, -1.260673, 1.570796, 1.865661],accel_mss,speed_ms,0,blend_radius_m)
  movel([0.302757, -0.630619, -2.813010, -1.268760, 1.570796, 1.873553],accel_mss,speed_ms,0,blend_radius_m)
  movel([0.306845, -0.626267, -2.813411, -1.272711, 1.570796, 1.877642],accel_mss,speed_ms,0,blend_radius_m)
  movel([0.310988, -0.622120, -2.813786, -1.276483, 1.570796, 1.881784],accel_mss,speed_ms,0,blend_radius_m)
  movel([0.315153, -0.618260, -2.814128, -1.280001, 1.570796, 1.885950],accel_mss,speed_ms,0,blend_radius_m)
  movel([0.319307, -0.614792, -2.814431, -1.283166, 1.570796, 1.890104],accel_mss,speed_ms,0,blend_radius_m)
  movel([0.323408, -0.611811, -2.814687, -1.285891, 1.570796, 1.894204],accel_mss,speed_ms,0,blend_radius_m)
  movel([0.327424, -0.609415, -2.814891, -1.288083, 1.570796, 1.898220],accel_mss,speed_ms,0,blend_radius_m)
  movel([0.335704, -0.605740, -2.815198, -1.291450, 1.570796, 1.906501],accel_mss,speed_ms,0,blend_radius_m)
  movel([0.338553, -0.604270, -2.815320, -1.292799, 1.570796, 1.909349],accel_mss,speed_ms,0,blend_radius_m)
  movel([0.341622, -0.602222, -2.815488, -1.294679, 1.570796, 1.912418],accel_mss,speed_ms,0,blend_radius_m)
  movel([0.344775, -0.599551, -2.815705, -1.297133, 1.570796, 1.915572],accel_mss,speed_ms,0,blend_radius_m)
  movel([0.347727, -0.596389, -2.815957, -1.300042, 1.570796, 1.918524],accel_mss,speed_ms,0,blend_radius_m)
  movel([0.349043, -0.594657, -2.816094, -1.301638, 1.570796, 1.919839],accel_mss,speed_ms,0,blend_radius_m)
  movel([0.350203, -0.592849, -2.816236, -1.303304, 1.570796, 1.920999],accel_mss,speed_ms,0,blend_radius_m)
  speed_ms = 0.005
  movel([0.350203, -0.587622, -2.809395, -1.315372, 1.570796, 1.920999],accel_mss,speed_ms,0,blend_radius_m)
  speed_ms = 0.040
  movel([0.368105, -0.554673, -2.811745, -1.345971, 1.570796, 1.938901],accel_mss,speed_ms,0,blend_radius_m)
  speed_ms = 0.005
  movel([0.368105, -0.559327, -2.818634, -1.334428, 1.570796, 1.938901],accel_mss,speed_ms,0,blend_radius_m)
  speed_ms = 0.025
  movel([0.368968, -0.559398, -2.818629, -1.334362, 1.570796, 1.939765],accel_mss,speed_ms,0,blend_radius_m)
  movel([0.368864, -0.560616, -2.818549, -1.333224, 1.570796, 1.939660],accel_mss,speed_ms,0,blend_radius_m)
  movel([0.368010, -0.562407, -2.818431, -1.331551, 1.570796, 1.938806],accel_mss,speed_ms,0,blend_radius_m)
  movel([0.366650, -0.564201, -2.818311, -1.329876, 1.570796, 1.937447],accel_mss,speed_ms,0,blend_radius_m)
  movel([0.365112, -0.565604, -2.818217, -1.328567, 1.570796, 1.935908],accel_mss,speed_ms,0,blend_radius_m)
  movel([0.363581, -0.566700, -2.818143, -1.327546, 1.570796, 1.934377],accel_mss,speed_ms,0,blend_radius_m)
  movel([0.360546, -0.568569, -2.818015, -1.325805, 1.570796, 1.931342],accel_mss,speed_ms,0,blend_radius_m)
  movel([0.358317, -0.570172, -2.817905, -1.324313, 1.570796, 1.929113],accel_mss,speed_ms,0,blend_radius_m)
  movel([0.356086, -0.572065, -2.817773, -1.322551, 1.570796, 1.926882],accel_mss,speed_ms,0,blend_radius_m)
  movel([0.351647, -0.576511, -2.817458, -1.318420, 1.570796, 1.922443],accel_mss,speed_ms,0,blend_radius_m)
  movel([0.347317, -0.581509, -2.817095, -1.313785, 1.570796, 1.918113],accel_mss,speed_ms,0,blend_radius_m)
  movel([0.343182, -0.586640, -2.816712, -1.309037, 1.570796, 1.913979],accel_mss,speed_ms,0,blend_radius_m)
  movel([0.342235, -0.587913, -2.816616, -1.307860, 1.570796, 1.913032],accel_mss,speed_ms,0,blend_radius_m)
  movel([0.341615, -0.589119, -2.816524, -1.306746, 1.570796, 1.912411],accel_mss,speed_ms,0,blend_radius_m)
  movel([0.341723, -0.589988, -2.816457, -1.305943, 1.570796, 1.912520],accel_mss,speed_ms,0,blend_radius_m)
  movel([0.342462, -0.590224, -2.816439, -1.305726, 1.570796, 1.913258],accel_mss,speed_ms,0,blend_radius_m)
  movel([0.344503, -0.590113, -2.816448, -1.305828, 1.570796, 1.915299],accel_mss,speed_ms,0,blend_radius_m)
  movel([0.346807, -0.589521, -2.816493, -1.306375, 1.570796, 1.917604],accel_mss,speed_ms,0,blend_radius_m)
  movel([0.349334, -0.588482, -2.816573, -1.307334, 1.570796, 1.920130],accel_mss,speed_ms,0,blend_radius_m)
  movel([0.352037, -0.587011, -2.816684, -1.308694, 1.570796, 1.922833],accel_mss,speed_ms,0,blend_radius_m)
  movel([0.354856, -0.585156, -2.816824, -1.310408, 1.570796, 1.925652],accel_mss,speed_ms,0,blend_radius_m)
  movel([0.357752, -0.582929, -2.816990, -1.312470, 1.570796, 1.928549],accel_mss,speed_ms,0,blend_radius_m)
  movel([0.360668, -0.580370, -2.817179, -1.314840, 1.570796, 1.931464],accel_mss,speed_ms,0,blend_radius_m)
  movel([0.363561, -0.577496, -2.817387, -1.317506, 1.570796, 1.934358],accel_mss,speed_ms,0,blend_radius_m)
  movel([0.362934, -0.579275, -2.817258, -1.315855, 1.570796, 1.933731],accel_mss,speed_ms,0,blend_radius_m)
  movel([0.363038, -0.580532, -2.817167, -1.314691, 1.570796, 1.933835],accel_mss,speed_ms,0,blend_radius_m)
  movel([0.363749, -0.581193, -2.817118, -1.314078, 1.570796, 1.934545],accel_mss,speed_ms,0,blend_radius_m)
  movel([0.364933, -0.581193, -2.817118, -1.314078, 1.570796, 1.935729],accel_mss,speed_ms,0,blend_radius_m)
  movel([0.366423, -0.580584, -2.817163, -1.314642, 1.570796, 1.937220],accel_mss,speed_ms,0,blend_radius_m)
  movel([0.368082, -0.579553, -2.817238, -1.315598, 1.570796, 1.938878],accel_mss,speed_ms,0,blend_radius_m)
  movel([0.371589, -0.576708, -2.817444, -1.318237, 1.570796, 1.942385],accel_mss,speed_ms,0,blend_radius_m)
  movel([0.376077, -0.572392, -2.817750, -1.322247, 1.570796, 1.946874],accel_mss,speed_ms,0,blend_radius_m)
  movel([0.380438, -0.567588, -2.818082, -1.326719, 1.570796, 1.951234],accel_mss,speed_ms,0,blend_radius_m)
  movel([0.384550, -0.562441, -2.818429, -1.331519, 1.570796, 1.955347],accel_mss,speed_ms,0,blend_radius_m)
  movel([0.388290, -0.557091, -2.818778, -1.336519, 1.570796, 1.959086],accel_mss,speed_ms,0,blend_radius_m)
  movel([0.389384, -0.555274, -2.818895, -1.338220, 1.570796, 1.960180],accel_mss,speed_ms,0,blend_radius_m)
  movel([0.389964, -0.553696, -2.818995, -1.339698, 1.570796, 1.960761],accel_mss,speed_ms,0,blend_radius_m)
  movel([0.389788, -0.552878, -2.819046, -1.340465, 1.570796, 1.960584],accel_mss,speed_ms,0,blend_radius_m)
  movel([0.389203, -0.552487, -2.819071, -1.340831, 1.570796, 1.959999],accel_mss,speed_ms,0,blend_radius_m)
  movel([0.386676, -0.551959, -2.819104, -1.341326, 1.570796, 1.957472],accel_mss,speed_ms,0,blend_radius_m)
  movel([0.381451, -0.551781, -2.819115, -1.341493, 1.570796, 1.952247],accel_mss,speed_ms,0,blend_radius_m)
  movel([0.379326, -0.550688, -2.819183, -1.342518, 1.570796, 1.950122],accel_mss,speed_ms,0,blend_radius_m)
  movel([0.384469, -0.544735, -2.819545, -1.348109, 1.570796, 1.955266],accel_mss,speed_ms,0,blend_radius_m)
  movel([0.387180, -0.542066, -2.819703, -1.350620, 1.570796, 1.957976],accel_mss,speed_ms,0,blend_radius_m)
  movel([0.389910, -0.539778, -2.819837, -1.352775, 1.570796, 1.960706],accel_mss,speed_ms,0,blend_radius_m)
  movel([0.391735, -0.538539, -2.819908, -1.353942, 1.570796, 1.962531],accel_mss,speed_ms,0,blend_radius_m)
  movel([0.393582, -0.537535, -2.819966, -1.354888, 1.570796, 1.964378],accel_mss,speed_ms,0,blend_radius_m)
  movel([0.396744, -0.536482, -2.820025, -1.355881, 1.570796, 1.967540],accel_mss,speed_ms,0,blend_radius_m)
  movel([0.398201, -0.536901, -2.820002, -1.355487, 1.570796, 1.968997],accel_mss,speed_ms,0,blend_radius_m)
  movel([0.398494, -0.537619, -2.819961, -1.354809, 1.570796, 1.969291],accel_mss,speed_ms,0,blend_radius_m)
  movel([0.398393, -0.538698, -2.819899, -1.353792, 1.570796, 1.969189],accel_mss,speed_ms,0,blend_radius_m)
  movel([0.397663, -0.540487, -2.819795, -1.352107, 1.570796, 1.968460],accel_mss,speed_ms,0,blend_radius_m)
  movel([0.396447, -0.542440, -2.819681, -1.350268, 1.570796, 1.967243],accel_mss,speed_ms,0,blend_radius_m)
  movel([0.393297, -0.546353, -2.819448, -1.346589, 1.570796, 1.964093],accel_mss,speed_ms,0,blend_radius_m)
  speed_ms = 0.005
  movel([0.393297, -0.541927, -2.812543, -1.357919, 1.570796, 1.964093],accel_mss,speed_ms,0,blend_radius_m)
  speed_ms = 0.040
  movel([0.440057, -0.416616, -2.817235, -1.478538, 1.570796, 2.010854],accel_mss,speed_ms,0,blend_radius_m)
  speed_ms = 0.005
  movel([0.440057, -0.418616, -2.824239, -1.469534, 1.570796, 2.010854],accel_mss,speed_ms,0,blend_radius_m)
  speed_ms = 0.025
  movel([0.442441, -0.416459, -2.824271, -1.471659, 1.570796, 2.013238],accel_mss,speed_ms,0,blend_radius_m)
  movel([0.444761, -0.414669, -2.824296, -1.473424, 1.570796, 2.015558],accel_mss,speed_ms,0,blend_radius_m)
  movel([0.446970, -0.413252, -2.824316, -1.474821, 1.570796, 2.017767],accel_mss,speed_ms,0,blend_radius_m)
  movel([0.450910, -0.411550, -2.824338, -1.476500, 1.570796, 2.021706],accel_mss,speed_ms,0,blend_radius_m)
  movel([0.452557, -0.411269, -2.824342, -1.476778, 1.570796, 2.023353],accel_mss,speed_ms,0,blend_radius_m)
  movel([0.455003, -0.411857, -2.824334, -1.476198, 1.570796, 2.025800],accel_mss,speed_ms,0,blend_radius_m)
  movel([0.456272, -0.413793, -2.824309, -1.474288, 1.570796, 2.027069],accel_mss,speed_ms,0,blend_radius_m)
  movel([0.456587, -0.416708, -2.824267, -1.471414, 1.570796, 2.027383],accel_mss,speed_ms,0,blend_radius_m)
  movel([0.456142, -0.420339, -2.824212, -1.467838, 1.570796, 2.026938],accel_mss,speed_ms,0,blend_radius_m)
  movel([0.455131, -0.424426, -2.824144, -1.463819, 1.570796, 2.025928],accel_mss,speed_ms,0,blend_radius_m)
  movel([0.452847, -0.431134, -2.824020, -1.457235, 1.570796, 2.023643],accel_mss,speed_ms,0,blend_radius_m)
  movel([0.449787, -0.438320, -2.823871, -1.450199, 1.570796, 2.020584],accel_mss,speed_ms,0,blend_radius_m)
  movel([0.446023, -0.445853, -2.823695, -1.442841, 1.570796, 2.016820],accel_mss,speed_ms,0,blend_radius_m)
  movel([0.437383, -0.460948, -2.823284, -1.428157, 1.570796, 2.008179],accel_mss,speed_ms,0,blend_radius_m)
  movel([0.435923, -0.464216, -2.823185, -1.424988, 1.570796, 2.006720],accel_mss,speed_ms,0,blend_radius_m)
  movel([0.435426, -0.466813, -2.823103, -1.422472, 1.570796, 2.006222],accel_mss,speed_ms,0,blend_radius_m)
  movel([0.435982, -0.468250, -2.823057, -1.421082, 1.570796, 2.006778],accel_mss,speed_ms,0,blend_radius_m)
  movel([0.437126, -0.469059, -2.823031, -1.420299, 1.570796, 2.007923],accel_mss,speed_ms,0,blend_radius_m)
  movel([0.438392, -0.469751, -2.823008, -1.419630, 1.570796, 2.009189],accel_mss,speed_ms,0,blend_radius_m)
  movel([0.439295, -0.470842, -2.822972, -1.418575, 1.570796, 2.010091],accel_mss,speed_ms,0,blend_radius_m)
  movel([0.439487, -0.472447, -2.822918, -1.417024, 1.570796, 2.010284],accel_mss,speed_ms,0,blend_radius_m)
  movel([0.439143, -0.474528, -2.822847, -1.415014, 1.570796, 2.009939],accel_mss,speed_ms,0,blend_radius_m)
  movel([0.437530, -0.479416, -2.822674, -1.410299, 1.570796, 2.008326],accel_mss,speed_ms,0,blend_radius_m)
  movel([0.434579, -0.486797, -2.822397, -1.403195, 1.570796, 2.005376],accel_mss,speed_ms,0,blend_radius_m)
  movel([0.431281, -0.494339, -2.822094, -1.395956, 1.570796, 2.002077],accel_mss,speed_ms,0,blend_radius_m)
  movel([0.427645, -0.502007, -2.821765, -1.388617, 1.570796, 1.998441],accel_mss,speed_ms,0,blend_radius_m)
  movel([0.423704, -0.509770, -2.821410, -1.381209, 1.570796, 1.994500],accel_mss,speed_ms,0,blend_radius_m)
  movel([0.419475, -0.517584, -2.821032, -1.373773, 1.570796, 1.990272],accel_mss,speed_ms,0,blend_radius_m)
  movel([0.414991, -0.525414, -2.820631, -1.366344, 1.570796, 1.985787],accel_mss,speed_ms,0,blend_radius_m)
  movel([0.410254, -0.533238, -2.820207, -1.358943, 1.570796, 1.981050],accel_mss,speed_ms,0,blend_radius_m)
  movel([0.405294, -0.541024, -2.819764, -1.351601, 1.570796, 1.976090],accel_mss,speed_ms,0,blend_radius_m)
  movel([0.401988, -0.545905, -2.819475, -1.347009, 1.570796, 1.972784],accel_mss,speed_ms,0,blend_radius_m)
  movel([0.398403, -0.550677, -2.819183, -1.342528, 1.570796, 1.969199],accel_mss,speed_ms,0,blend_radius_m)
  movel([0.394613, -0.554973, -2.818914, -1.338502, 1.570796, 1.965409],accel_mss,speed_ms,0,blend_radius_m)
  movel([0.392667, -0.556817, -2.818796, -1.336776, 1.570796, 1.963463],accel_mss,speed_ms,0,blend_radius_m)
  movel([0.390691, -0.558412, -2.818693, -1.335284, 1.570796, 1.961488],accel_mss,speed_ms,0,blend_radius_m)
  speed_ms = 0.005
  movel([0.390691, -0.553773, -2.811803, -1.346812, 1.570796, 1.961488],accel_mss,speed_ms,0,blend_radius_m)
  speed_ms = 0.040
  movel([0.379771, -0.567139, -2.810905, -1.334345, 1.570796, 1.950568],accel_mss,speed_ms,0,blend_radius_m)
  speed_ms = 0.005
  movel([0.379771, -0.572014, -2.817776, -1.322599, 1.570796, 1.950568],accel_mss,speed_ms,0,blend_radius_m)
  speed_ms = 0.025
  movel([0.379949, -0.573051, -2.817704, -1.321635, 1.570796, 1.950745],accel_mss,speed_ms,0,blend_radius_m)
  movel([0.379468, -0.574621, -2.817593, -1.320175, 1.570796, 1.950264],accel_mss,speed_ms,0,blend_radius_m)
  movel([0.378499, -0.576458, -2.817462, -1.318470, 1.570796, 1.949295],accel_mss,speed_ms,0,blend_radius_m)
  movel([0.377199, -0.578293, -2.817330, -1.316766, 1.570796, 1.947995],accel_mss,speed_ms,0,blend_radius_m)
  movel([0.375432, -0.580154, -2.817194, -1.315040, 1.570796, 1.946228],accel_mss,speed_ms,0,blend_radius_m)
  movel([0.373657, -0.581632, -2.817086, -1.313671, 1.570796, 1.944453],accel_mss,speed_ms,0,blend_radius_m)
  movel([0.371926, -0.583016, -2.816984, -1.312389, 1.570796, 1.942722],accel_mss,speed_ms,0,blend_radius_m)
  movel([0.370313, -0.584595, -2.816866, -1.310927, 1.570796, 1.941109],accel_mss,speed_ms,0,blend_radius_m)
  movel([0.368536, -0.587266, -2.816665, -1.308458, 1.570796, 1.939332],accel_mss,speed_ms,0,blend_radius_m)
  movel([0.367706, -0.588655, -2.816559, -1.307175, 1.570796, 1.938503],accel_mss,speed_ms,0,blend_radius_m)
  movel([0.366616, -0.590129, -2.816446, -1.305814, 1.570796, 1.937412],accel_mss,speed_ms,0,blend_radius_m)
  movel([0.363281, -0.593784, -2.816163, -1.302443, 1.570796, 1.934078],accel_mss,speed_ms,0,blend_radius_m)
  movel([0.359964, -0.596927, -2.815915, -1.299547, 1.570796, 1.930761],accel_mss,speed_ms,0,blend_radius_m)
  movel([0.356635, -0.599637, -2.815698, -1.297054, 1.570796, 1.927431],accel_mss,speed_ms,0,blend_radius_m)
  movel([0.353259, -0.602019, -2.815505, -1.294865, 1.570796, 1.924055],accel_mss,speed_ms,0,blend_radius_m)
  movel([0.355034, -0.600604, -2.815620, -1.296165, 1.570796, 1.925830],accel_mss,speed_ms,0,blend_radius_m)
  movel([0.356757, -0.599464, -2.815712, -1.297213, 1.570796, 1.927553],accel_mss,speed_ms,0,blend_radius_m)
  movel([0.358252, -0.598961, -2.815752, -1.297676, 1.570796, 1.929048],accel_mss,speed_ms,0,blend_radius_m)
  movel([0.359104, -0.599449, -2.815713, -1.297227, 1.570796, 1.929901],accel_mss,speed_ms,0,blend_radius_m)
  movel([0.358949, -0.600950, -2.815591, -1.295847, 1.570796, 1.929745],accel_mss,speed_ms,0,blend_radius_m)
  movel([0.358015, -0.602921, -2.815431, -1.294037, 1.570796, 1.928811],accel_mss,speed_ms,0,blend_radius_m)
  movel([0.356611, -0.604918, -2.815267, -1.292204, 1.570796, 1.927407],accel_mss,speed_ms,0,blend_radius_m)
  movel([0.352353, -0.609671, -2.814869, -1.287849, 1.570796, 1.923149],accel_mss,speed_ms,0,blend_radius_m)
  movel([0.349628, -0.612299, -2.814646, -1.285445, 1.570796, 1.920424],accel_mss,speed_ms,0,blend_radius_m)
  movel([0.346894, -0.614652, -2.814443, -1.283294, 1.570796, 1.917690],accel_mss,speed_ms,0,blend_radius_m)
  movel([0.344176, -0.616702, -2.814265, -1.281422, 1.570796, 1.914972],accel_mss,speed_ms,0,blend_radius_m)
  movel([0.347204, -0.614806, -2.814430, -1.283153, 1.570796, 1.918001],accel_mss,speed_ms,0,blend_radius_m)
  movel([0.350417, -0.612444, -2.814633, -1.285312, 1.570796, 1.921214],accel_mss,speed_ms,0,blend_radius_m)
  movel([0.353558, -0.610198, -2.814825, -1.287366, 1.570796, 1.924354],accel_mss,speed_ms,0,blend_radius_m)
  movel([0.356373, -0.608624, -2.814957, -1.288807, 1.570796, 1.927169],accel_mss,speed_ms,0,blend_radius_m)
  movel([0.357104, -0.608552, -2.814964, -1.288874, 1.570796, 1.927900],accel_mss,speed_ms,0,blend_radius_m)
  movel([0.357042, -0.609160, -2.814912, -1.288317, 1.570796, 1.927838],accel_mss,speed_ms,0,blend_radius_m)
  movel([0.355138, -0.612416, -2.814636, -1.285337, 1.570796, 1.925934],accel_mss,speed_ms,0,blend_radius_m)
  movel([0.353460, -0.614779, -2.814432, -1.283177, 1.570796, 1.924257],accel_mss,speed_ms,0,blend_radius_m)
  movel([0.351629, -0.617048, -2.814235, -1.281106, 1.570796, 1.922426],accel_mss,speed_ms,0,blend_radius_m)
  movel([0.349693, -0.619160, -2.814049, -1.279180, 1.570796, 1.920490],accel_mss,speed_ms,0,blend_radius_m)
  movel([0.350644, -0.618339, -2.814121, -1.279929, 1.570796, 1.921441],accel_mss,speed_ms,0,blend_radius_m)
  movel([0.351670, -0.617715, -2.814176, -1.280498, 1.570796, 1.922466],accel_mss,speed_ms,0,blend_radius_m)
  movel([0.353820, -0.617011, -2.814238, -1.281140, 1.570796, 1.924616],accel_mss,speed_ms,0,blend_radius_m)
  movel([0.355869, -0.616979, -2.814241, -1.281169, 1.570796, 1.926665],accel_mss,speed_ms,0,blend_radius_m)
  movel([0.357562, -0.617534, -2.814192, -1.280663, 1.570796, 1.928358],accel_mss,speed_ms,0,blend_radius_m)
  movel([0.358648, -0.618587, -2.814100, -1.279702, 1.570796, 1.929444],accel_mss,speed_ms,0,blend_radius_m)
  movel([0.358876, -0.620042, -2.813971, -1.278376, 1.570796, 1.929673],accel_mss,speed_ms,0,blend_radius_m)
  movel([0.358591, -0.620890, -2.813896, -1.277603, 1.570796, 1.929388],accel_mss,speed_ms,0,blend_radius_m)
  movel([0.357999, -0.621800, -2.813814, -1.276774, 1.570796, 1.928795],accel_mss,speed_ms,0,blend_radius_m)
  movel([0.357072, -0.622771, -2.813727, -1.275890, 1.570796, 1.927869],accel_mss,speed_ms,0,blend_radius_m)
  movel([0.355773, -0.623782, -2.813636, -1.274970, 1.570796, 1.926569],accel_mss,speed_ms,0,blend_radius_m)
  movel([0.354385, -0.624511, -2.813571, -1.274307, 1.570796, 1.925181],accel_mss,speed_ms,0,blend_radius_m)
  movel([0.349446, -0.625337, -2.813496, -1.273556, 1.570796, 1.920242],accel_mss,speed_ms,0,blend_radius_m)
  movel([0.347504, -0.625788, -2.813455, -1.273147, 1.570796, 1.918301],accel_mss,speed_ms,0,blend_radius_m)
  movel([0.345366, -0.626694, -2.813372, -1.272323, 1.570796, 1.916163],accel_mss,speed_ms,0,blend_radius_m)
  movel([0.341503, -0.629264, -2.813136, -1.269989, 1.570796, 1.912300],accel_mss,speed_ms,0,blend_radius_m)
  movel([0.337576, -0.632126, -2.812870, -1.267393, 1.570796, 1.908372],accel_mss,speed_ms,0,blend_radius_m)
  movel([0.335660, -0.633229, -2.812767, -1.266394, 1.570796, 1.906456],accel_mss,speed_ms,0,blend_radius_m)
  movel([0.333925, -0.633855, -2.812708, -1.265826, 1.570796, 1.904721],accel_mss,speed_ms,0,blend_radius_m)
  movel([0.332602, -0.633818, -2.812711, -1.265860, 1.570796, 1.903398],accel_mss,speed_ms,0,blend_radius_m)
  movel([0.331912, -0.632941, -2.812794, -1.266655, 1.570796, 1.902709],accel_mss,speed_ms,0,blend_radius_m)
  movel([0.333990, -0.630244, -2.813045, -1.269100, 1.570796, 1.904787],accel_mss,speed_ms,0,blend_radius_m)
  movel([0.336211, -0.627669, -2.813283, -1.271437, 1.570796, 1.907007],accel_mss,speed_ms,0,blend_radius_m)
  speed_ms = 0.005
  movel([0.336211, -0.621877, -2.806500, -1.284012, 1.570796, 1.907007],accel_mss,speed_ms,0,blend_radius_m)
  speed_ms = 0.040
  movel([0.351549, -0.631195, -2.805631, -1.275563, 1.570796, 1.922345],accel_mss,speed_ms,0,blend_radius_m)
  speed_ms = 0.005
  movel([0.351549, -0.637136, -2.812396, -1.262857, 1.570796, 1.922345],accel_mss,speed_ms,0,blend_radius_m)
  speed_ms = 0.025
  movel([0.353017, -0.635212, -2.812579, -1.264598, 1.570796, 1.923813],accel_mss,speed_ms,0,blend_radius_m)
  movel([0.354736, -0.633739, -2.812719, -1.265931, 1.570796, 1.925532],accel_mss,speed_ms,0,blend_radius_m)
  movel([0.356426, -0.632842, -2.812803, -1.266744, 1.570796, 1.927223],accel_mss,speed_ms,0,blend_radius_m)
  movel([0.357799, -0.632658, -2.812820, -1.266911, 1.570796, 1.928595],accel_mss,speed_ms,0,blend_radius_m)
  movel([0.358713, -0.633135, -2.812775, -1.266479, 1.570796, 1.929509],accel_mss,speed_ms,0,blend_radius_m)
  movel([0.359289, -0.634035, -2.812691, -1.265663, 1.570796, 1.930085],accel_mss,speed_ms,0,blend_radius_m)
  movel([0.359851, -0.636501, -2.812457, -1.263431, 1.570796, 1.930648],accel_mss,speed_ms,0,blend_radius_m)
  movel([0.361230, -0.634153, -2.812680, -1.265557, 1.570796, 1.932027],accel_mss,speed_ms,0,blend_radius_m)
  movel([0.362162, -0.631897, -2.812891, -1.267600, 1.570796, 1.932958],accel_mss,speed_ms,0,blend_radius_m)
  movel([0.362570, -0.629931, -2.813074, -1.269384, 1.570796, 1.933367],accel_mss,speed_ms,0,blend_radius_m)
  movel([0.362409, -0.628414, -2.813214, -1.270761, 1.570796, 1.933205],accel_mss,speed_ms,0,blend_radius_m)
  movel([0.363247, -0.628833, -2.813176, -1.270380, 1.570796, 1.934044],accel_mss,speed_ms,0,blend_radius_m)
  movel([0.363803, -0.629584, -2.813106, -1.269698, 1.570796, 1.934599],accel_mss,speed_ms,0,blend_radius_m)
  movel([0.364218, -0.631851, -2.812896, -1.267642, 1.570796, 1.935014],accel_mss,speed_ms,0,blend_radius_m)
  movel([0.363986, -0.634780, -2.812620, -1.264989, 1.570796, 1.934783],accel_mss,speed_ms,0,blend_radius_m)
  movel([0.363403, -0.637970, -2.812316, -1.262103, 1.570796, 1.934200],accel_mss,speed_ms,0,blend_radius_m)
  movel([0.362304, -0.641694, -2.811956, -1.258739, 1.570796, 1.933101],accel_mss,speed_ms,0,blend_radius_m)
  movel([0.360800, -0.645415, -2.811591, -1.255384, 1.570796, 1.931596],accel_mss,speed_ms,0,blend_radius_m)
  movel([0.359255, -0.649085, -2.811224, -1.252079, 1.570796, 1.930051],accel_mss,speed_ms,0,blend_radius_m)
  movel([0.358028, -0.652673, -2.810861, -1.248855, 1.570796, 1.928824],accel_mss,speed_ms,0,blend_radius_m)
  movel([0.357067, -0.651094, -2.811022, -1.250273, 1.570796, 1.927863],accel_mss,speed_ms,0,blend_radius_m)
  movel([0.355532, -0.650238, -2.811108, -1.251043, 1.570796, 1.926329],accel_mss,speed_ms,0,blend_radius_m)
  movel([0.353464, -0.650179, -2.811114, -1.251096, 1.570796, 1.924261],accel_mss,speed_ms,0,blend_radius_m)
  movel([0.350894, -0.650994, -2.811032, -1.250363, 1.570796, 1.921690],accel_mss,speed_ms,0,blend_radius_m)
  speed_ms = 0.005
  movel([0.350894, -0.644841, -2.804293, -1.263255, 1.570796, 1.921690],accel_mss,speed_ms,0,blend_radius_m)
  speed_ms = 0.040
  movel([0.352138, -0.654209, -2.803329, -1.254851, 1.570796, 1.922935],accel_mss,speed_ms,0,blend_radius_m)
  speed_ms = 0.005
  movel([0.352138, -0.660504, -2.810049, -1.241836, 1.570796, 1.922935],accel_mss,speed_ms,0,blend_radius_m)
  speed_ms = 0.025
  movel([0.351964, -0.664554, -2.809619, -1.238216, 1.570796, 1.922760],accel_mss,speed_ms,0,blend_radius_m)
  movel([0.352428, -0.668043, -2.809243, -1.235102, 1.570796, 1.923224],accel_mss,speed_ms,0,blend_radius_m)
  movel([0.353764, -0.670550, -2.808970, -1.232869, 1.570796, 1.924560],accel_mss,speed_ms,0,blend_radius_m)
  movel([0.354836, -0.671301, -2.808888, -1.232200, 1.570796, 1.925632],accel_mss,speed_ms,0,blend_radius_m)
  movel([0.356219, -0.671650, -2.808849, -1.231890, 1.570796, 1.927016],accel_mss,speed_ms,0,blend_radius_m)
  movel([0.358558, -0.671408, -2.808876, -1.232105, 1.570796, 1.929355],accel_mss,speed_ms,0,blend_radius_m)
  movel([0.361206, -0.670458, -2.808980, -1.232951, 1.570796, 1.932002],accel_mss,speed_ms,0,blend_radius_m)
  movel([0.364101, -0.668960, -2.809144, -1.234285, 1.570796, 1.934897],accel_mss,speed_ms,0,blend_radius_m)
  movel([0.367174, -0.667079, -2.809348, -1.235962, 1.570796, 1.937971],accel_mss,speed_ms,0,blend_radius_m)
  movel([0.373586, -0.662812, -2.809805, -1.239772, 1.570796, 1.944382],accel_mss,speed_ms,0,blend_radius_m)
  movel([0.379870, -0.658991, -2.810208, -1.243190, 1.570796, 1.950666],accel_mss,speed_ms,0,blend_radius_m)
  movel([0.383258, -0.657485, -2.810365, -1.244539, 1.570796, 1.954054],accel_mss,speed_ms,0,blend_radius_m)
  movel([0.386363, -0.656638, -2.810453, -1.245298, 1.570796, 1.957160],accel_mss,speed_ms,0,blend_radius_m)
  movel([0.389136, -0.656435, -2.810474, -1.245480, 1.570796, 1.959932],accel_mss,speed_ms,0,blend_radius_m)
  movel([0.391521, -0.656870, -2.810429, -1.245090, 1.570796, 1.962317],accel_mss,speed_ms,0,blend_radius_m)
  movel([0.393479, -0.657914, -2.810321, -1.244154, 1.570796, 1.964275],accel_mss,speed_ms,0,blend_radius_m)
  movel([0.394959, -0.659557, -2.810149, -1.242683, 1.570796, 1.965755],accel_mss,speed_ms,0,blend_radius_m)
  movel([0.395914, -0.661777, -2.809915, -1.240697, 1.570796, 1.966710],accel_mss,speed_ms,0,blend_radius_m)
  movel([0.396312, -0.664541, -2.809621, -1.238227, 1.570796, 1.967108],accel_mss,speed_ms,0,blend_radius_m)
  speed_ms = 0.005
  movel([0.396312, -0.658186, -2.802909, -1.251294, 1.570796, 1.967108],accel_mss,speed_ms,0,blend_radius_m)
  speed_ms = 0.040
  movel([0.345905, -0.626699, -2.806055, -1.279635, 1.570796, 1.916701],accel_mss,speed_ms,0,blend_radius_m)
  speed_ms = 0.005
  movel([0.345905, -0.632568, -2.812829, -1.266992, 1.570796, 1.916701],accel_mss,speed_ms,0,blend_radius_m)
  speed_ms = 0.025
  movel([0.347293, -0.632878, -2.812800, -1.266712, 1.570796, 1.918089],accel_mss,speed_ms,0,blend_radius_m)
  movel([0.348210, -0.633782, -2.812714, -1.265893, 1.570796, 1.919007],accel_mss,speed_ms,0,blend_radius_m)
  movel([0.348304, -0.634634, -2.812634, -1.265121, 1.570796, 1.919100],accel_mss,speed_ms,0,blend_radius_m)
  movel([0.348070, -0.635744, -2.812529, -1.264116, 1.570796, 1.918866],accel_mss,speed_ms,0,blend_radius_m)
  movel([0.347517, -0.636989, -2.812410, -1.262990, 1.570796, 1.918313],accel_mss,speed_ms,0,blend_radius_m)
  movel([0.346644, -0.638247, -2.812290, -1.261852, 1.570796, 1.917440],accel_mss,speed_ms,0,blend_radius_m)
  movel([0.344727, -0.640332, -2.812089, -1.259969, 1.570796, 1.915523],accel_mss,speed_ms,0,blend_radius_m)
  movel([0.343988, -0.641521, -2.811973, -1.258895, 1.570796, 1.914784],accel_mss,speed_ms,0,blend_radius_m)
  movel([0.343592, -0.642641, -2.811864, -1.257884, 1.570796, 1.914388],accel_mss,speed_ms,0,blend_radius_m)
  movel([0.343551, -0.644491, -2.811682, -1.256216, 1.570796, 1.914347],accel_mss,speed_ms,0,blend_radius_m)
  movel([0.344108, -0.646100, -2.811523, -1.254767, 1.570796, 1.914905],accel_mss,speed_ms,0,blend_radius_m)
  movel([0.345022, -0.647314, -2.811402, -1.253673, 1.570796, 1.915818],accel_mss,speed_ms,0,blend_radius_m)
  movel([0.346266, -0.648131, -2.811320, -1.252938, 1.570796, 1.917062],accel_mss,speed_ms,0,blend_radius_m)
  movel([0.347814, -0.648518, -2.811281, -1.252590, 1.570796, 1.918611],accel_mss,speed_ms,0,blend_radius_m)
  movel([0.346143, -0.651177, -2.811013, -1.250199, 1.570796, 1.916940],accel_mss,speed_ms,0,blend_radius_m)
  movel([0.344813, -0.653762, -2.810750, -1.247877, 1.570796, 1.915609],accel_mss,speed_ms,0,blend_radius_m)
  movel([0.343783, -0.656270, -2.810491, -1.245628, 1.570796, 1.914580],accel_mss,speed_ms,0,blend_radius_m)
  movel([0.343015, -0.658691, -2.810240, -1.243459, 1.570796, 1.913812],accel_mss,speed_ms,0,blend_radius_m)
  movel([0.342123, -0.663236, -2.809760, -1.239393, 1.570796, 1.912920],accel_mss,speed_ms,0,blend_radius_m)
  movel([0.341863, -0.667326, -2.809321, -1.235742, 1.570796, 1.912659],accel_mss,speed_ms,0,blend_radius_m)
  movel([0.341691, -0.671213, -2.808897, -1.232278, 1.570796, 1.912487],accel_mss,speed_ms,0,blend_radius_m)
  movel([0.341301, -0.673346, -2.808662, -1.230381, 1.570796, 1.912097],accel_mss,speed_ms,0,blend_radius_m)
  movel([0.340520, -0.675694, -2.808401, -1.228294, 1.570796, 1.911316],accel_mss,speed_ms,0,blend_radius_m)
  movel([0.339172, -0.678276, -2.808111, -1.226002, 1.570796, 1.909969],accel_mss,speed_ms,0,blend_radius_m)
  movel([0.337350, -0.680806, -2.807824, -1.223759, 1.570796, 1.908147],accel_mss,speed_ms,0,blend_radius_m)
  movel([0.335304, -0.682889, -2.807585, -1.221914, 1.570796, 1.906101],accel_mss,speed_ms,0,blend_radius_m)
  movel([0.333296, -0.684121, -2.807443, -1.220825, 1.570796, 1.904092],accel_mss,speed_ms,0,blend_radius_m)
  movel([0.333851, -0.685420, -2.807293, -1.219676, 1.570796, 1.904647],accel_mss,speed_ms,0,blend_radius_m)
  movel([0.334133, -0.688796, -2.806899, -1.216694, 1.570796, 1.904930],accel_mss,speed_ms,0,blend_radius_m)
  movel([0.333871, -0.690805, -2.806662, -1.214922, 1.570796, 1.904667],accel_mss,speed_ms,0,blend_radius_m)
  movel([0.332594, -0.695273, -2.806129, -1.210987, 1.570796, 1.903390],accel_mss,speed_ms,0,blend_radius_m)
  movel([0.331591, -0.697661, -2.805840, -1.208888, 1.570796, 1.902387],accel_mss,speed_ms,0,blend_radius_m)
  movel([0.330351, -0.700112, -2.805541, -1.206736, 1.570796, 1.901147],accel_mss,speed_ms,0,blend_radius_m)
  speed_ms = 0.005
  movel([0.330351, -0.693251, -2.798906, -1.220231, 1.570796, 1.901147],accel_mss,speed_ms,0,blend_radius_m)
  speed_ms = 0.040
  movel([0.320831, -0.697283, -2.798411, -1.216694, 1.570796, 1.891628],accel_mss,speed_ms,0,blend_radius_m)
  speed_ms = 0.005
  movel([0.320831, -0.704199, -2.805037, -1.203153, 1.570796, 1.891628],accel_mss,speed_ms,0,blend_radius_m)
  speed_ms = 0.025
  movel([0.323413, -0.720922, -2.802895, -1.188572, 1.570796, 1.894209],accel_mss,speed_ms,0,blend_radius_m)
  movel([0.323461, -0.723179, -2.802596, -1.186614, 1.570796, 1.894258],accel_mss,speed_ms,0,blend_radius_m)
  movel([0.323113, -0.724501, -2.802420, -1.185468, 1.570796, 1.893909],accel_mss,speed_ms,0,blend_radius_m)
  movel([0.322352, -0.725941, -2.802227, -1.184221, 1.570796, 1.893148],accel_mss,speed_ms,0,blend_radius_m)
  movel([0.320056, -0.728986, -2.801816, -1.181587, 1.570796, 1.890852],accel_mss,speed_ms,0,blend_radius_m)
  movel([0.319501, -0.730490, -2.801612, -1.180287, 1.570796, 1.890297],accel_mss,speed_ms,0,blend_radius_m)
  movel([0.319482, -0.731720, -2.801444, -1.179225, 1.570796, 1.890279],accel_mss,speed_ms,0,blend_radius_m)
  movel([0.320112, -0.733196, -2.801241, -1.177952, 1.570796, 1.890908],accel_mss,speed_ms,0,blend_radius_m)
  movel([0.321291, -0.734151, -2.801110, -1.177129, 1.570796, 1.892088],accel_mss,speed_ms,0,blend_radius_m)
  movel([0.323990, -0.735536, -2.800918, -1.175935, 1.570796, 1.894786],accel_mss,speed_ms,0,blend_radius_m)
  movel([0.325329, -0.736999, -2.800715, -1.174676, 1.570796, 1.896125],accel_mss,speed_ms,0,blend_radius_m)
  movel([0.326698, -0.739636, -2.800345, -1.172408, 1.570796, 1.897494],accel_mss,speed_ms,0,blend_radius_m)
  movel([0.326968, -0.741136, -2.800134, -1.171119, 1.570796, 1.897764],accel_mss,speed_ms,0,blend_radius_m)
  movel([0.326754, -0.742610, -2.799925, -1.169854, 1.570796, 1.897550],accel_mss,speed_ms,0,blend_radius_m)
  movel([0.326410, -0.743302, -2.799827, -1.169261, 1.570796, 1.897207],accel_mss,speed_ms,0,blend_radius_m)
  movel([0.325881, -0.743946, -2.799735, -1.168708, 1.570796, 1.896678],accel_mss,speed_ms,0,blend_radius_m)
  movel([0.324184, -0.745054, -2.799576, -1.167758, 1.570796, 1.894981],accel_mss,speed_ms,0,blend_radius_m)
  movel([0.324146, -0.746517, -2.799366, -1.166505, 1.570796, 1.894943],accel_mss,speed_ms,0,blend_radius_m)
  movel([0.324547, -0.747842, -2.799175, -1.165372, 1.570796, 1.895344],accel_mss,speed_ms,0,blend_radius_m)
  movel([0.326252, -0.750067, -2.798852, -1.163469, 1.570796, 1.897049],accel_mss,speed_ms,0,blend_radius_m)
  movel([0.330428, -0.752907, -2.798437, -1.161045, 1.570796, 1.901225],accel_mss,speed_ms,0,blend_radius_m)
  movel([0.332973, -0.753684, -2.798323, -1.160382, 1.570796, 1.903769],accel_mss,speed_ms,0,blend_radius_m)
  movel([0.335888, -0.754127, -2.798257, -1.160005, 1.570796, 1.906684],accel_mss,speed_ms,0,blend_radius_m)
  movel([0.338411, -0.755040, -2.798122, -1.159226, 1.570796, 1.909207],accel_mss,speed_ms,0,blend_radius_m)
  movel([0.339288, -0.755918, -2.797992, -1.158478, 1.570796, 1.910085],accel_mss,speed_ms,0,blend_radius_m)
  movel([0.339784, -0.757209, -2.797800, -1.157380, 1.570796, 1.910580],accel_mss,speed_ms,0,blend_radius_m)
  movel([0.339779, -0.758105, -2.797666, -1.156618, 1.570796, 1.910575],accel_mss,speed_ms,0,blend_radius_m)
  movel([0.339496, -0.759170, -2.797507, -1.155712, 1.570796, 1.910293],accel_mss,speed_ms,0,blend_radius_m)
  movel([0.338944, -0.760213, -2.797350, -1.154825, 1.570796, 1.909740],accel_mss,speed_ms,0,blend_radius_m)
  movel([0.338115, -0.761041, -2.797225, -1.154123, 1.570796, 1.908911],accel_mss,speed_ms,0,blend_radius_m)
  movel([0.336844, -0.761370, -2.797176, -1.153843, 1.570796, 1.907640],accel_mss,speed_ms,0,blend_radius_m)
  movel([0.331845, -0.760698, -2.797277, -1.154414, 1.570796, 1.902641],accel_mss,speed_ms,0,blend_radius_m)
  movel([0.327463, -0.759082, -2.797520, -1.155787, 1.570796, 1.898259],accel_mss,speed_ms,0,blend_radius_m)
  movel([0.326911, -0.760259, -2.797343, -1.154787, 1.570796, 1.897708],accel_mss,speed_ms,0,blend_radius_m)
  movel([0.326609, -0.761345, -2.797180, -1.153864, 1.570796, 1.897405],accel_mss,speed_ms,0,blend_radius_m)
  movel([0.326653, -0.763259, -2.796889, -1.152240, 1.570796, 1.897450],accel_mss,speed_ms,0,blend_radius_m)
  movel([0.327394, -0.764849, -2.796647, -1.150893, 1.570796, 1.898190],accel_mss,speed_ms,0,blend_radius_m)
  movel([0.328616, -0.766167, -2.796445, -1.149777, 1.570796, 1.899412],accel_mss,speed_ms,0,blend_radius_m)
  movel([0.331744, -0.768072, -2.796152, -1.148165, 1.570796, 1.902540],accel_mss,speed_ms,0,blend_radius_m)
  movel([0.334451, -0.769215, -2.795975, -1.147198, 1.570796, 1.905247],accel_mss,speed_ms,0,blend_radius_m)
  movel([0.335324, -0.769810, -2.795883, -1.146696, 1.570796, 1.906121],accel_mss,speed_ms,0,blend_radius_m)
  movel([0.335511, -0.770343, -2.795800, -1.146246, 1.570796, 1.906307],accel_mss,speed_ms,0,blend_radius_m)
  movel([0.335387, -0.771111, -2.795681, -1.145598, 1.570796, 1.906183],accel_mss,speed_ms,0,blend_radius_m)
  movel([0.334923, -0.772065, -2.795532, -1.144792, 1.570796, 1.905720],accel_mss,speed_ms,0,blend_radius_m)
  movel([0.334354, -0.772756, -2.795423, -1.144209, 1.570796, 1.905150],accel_mss,speed_ms,0,blend_radius_m)
  movel([0.333034, -0.773619, -2.795288, -1.143482, 1.570796, 1.903831],accel_mss,speed_ms,0,blend_radius_m)
  movel([0.331203, -0.774628, -2.795129, -1.142632, 1.570796, 1.901999],accel_mss,speed_ms,0,blend_radius_m)
  movel([0.330790, -0.775155, -2.795046, -1.142188, 1.570796, 1.901586],accel_mss,speed_ms,0,blend_radius_m)
  movel([0.330501, -0.775943, -2.794921, -1.141525, 1.570796, 1.901297],accel_mss,speed_ms,0,blend_radius_m)
  movel([0.330491, -0.776663, -2.794807, -1.140918, 1.570796, 1.901287],accel_mss,speed_ms,0,blend_radius_m)
  movel([0.331058, -0.777890, -2.794612, -1.139887, 1.570796, 1.901854],accel_mss,speed_ms,0,blend_radius_m)
  movel([0.332754, -0.779530, -2.794350, -1.138509, 1.570796, 1.903551],accel_mss,speed_ms,0,blend_radius_m)
  movel([0.340812, -0.785407, -2.793400, -1.133581, 1.570796, 1.911608],accel_mss,speed_ms,0,blend_radius_m)
  movel([0.341451, -0.786207, -2.793270, -1.132912, 1.570796, 1.912247],accel_mss,speed_ms,0,blend_radius_m)
  movel([0.341793, -0.787306, -2.793090, -1.131993, 1.570796, 1.912589],accel_mss,speed_ms,0,blend_radius_m)
  movel([0.341637, -0.788664, -2.792866, -1.130858, 1.570796, 1.912433],accel_mss,speed_ms,0,blend_radius_m)
  movel([0.340781, -0.790231, -2.792608, -1.129551, 1.570796, 1.911578],accel_mss,speed_ms,0,blend_radius_m)
  movel([0.339541, -0.791437, -2.792408, -1.128545, 1.570796, 1.910338],accel_mss,speed_ms,0,blend_radius_m)
  movel([0.338270, -0.792048, -2.792306, -1.128035, 1.570796, 1.909067],accel_mss,speed_ms,0,blend_radius_m)
